(* IEC 61131-3 sources: daoli-st-library/DL_Process (part 48) *)

(* ---- FB_DL_RecipeSwitchHandover.st ---- *)
(*
  Name        : FB_DL_RecipeSwitchHandover
  Category    : DL_Process
  Version     : 1.0.0
  Purpose     : 配方切换交接编排：旧配方排空确认 → 参数装载复核（校验和整数直比）→ 新配方放行三相时序，各相独立超时故障码，中止命令相边界停下；/ Recipe switch handover orchestration: drain confirm, load recheck by integer checksum compare, release three-phase sequence with per-phase timeout fault codes and abort at phase boundary
  溯源        : 借 packml/isa88 的配方切换/批次编排组织，clean-room 实现
  Boundary    : ① 三相（排空确认/装载复核/放行）各自 TON 断输入归零 + 相超时独立锁存故障码（R40/R44）；
                ② 装载复核 = 参数集校验和整数直比，不符不放行不半装载（锁存故障至复位沿）；
                ③ 切换中收到中止命令 → 当前相边界停下（不回滚已装载段，eHold 相状态可查，信息级成因）；
                ④ 放行前复核旧配方累计量已清零反馈（幂等放行），未清零不放行（锁存故障）；
                ⑤ 命令优先级：中止 > 放行 > 装载，低优先命令直接丢弃不排队（放行仅放行相生效，装载仅空闲相受理）。
*)
TYPE E_DL_RshState :
(
    eIdle    := 0,                           (* 空闲（可受理装载命令） / Idle *)
    eDrain   := 10,                          (* 旧配方排空确认相 / Drain confirm *)
    eLoadChk := 20,                          (* 参数装载复核相 / Load recheck *)
    eRelease := 30,                          (* 新配方放行相 / Release *)
    eHold    := 40,                          (* 中止驻留相（状态可查） / Abort hold *)
    eFault   := 90                           (* 故障锁存相 / Fault latched *)
);
END_TYPE

TYPE E_DL_RshCause :
(
    eNone      := 0,                         (* 无成因 / No cause *)
    eCfgIllegal:= 1,                        (* 组态非法：相超时/周期域越界 / Illegal config *)
    eDrainTo   := 2,                        (* 排空相超时（独立码，边界①） / Drain timeout *)
    eLoadTo    := 3,                        (* 装载复核相超时（独立码） / Load recheck timeout *)
    eRelTo     := 4,                        (* 放行相超时（独立码） / Release timeout *)
    eChkMis    := 5,                        (* 校验和不符（不放行不半装载，边界②） / Checksum mismatch *)
    eAccNotClr := 6,                         (* 旧累计量未清零（不放行，边界④） / Accumulator not cleared *)
    eAbort     := 7,                        (* 中止驻留（信息级，边界③） / Abort hold, info level *)
    ePhaseBad  := 8                         (* 非法相位兜底 / Illegal phase fallback *)
);
END_TYPE

FUNCTION_BLOCK FB_DL_RecipeSwitchHandover
VAR_INPUT
    bCmdLoad : BOOL := FALSE;                (* 装载命令（仅空闲相受理，低优先丢弃）[-] / Load command *)
    bCmdRelease: BOOL := FALSE;              (* 放行命令（仅放行相复核生效）[-] / Release command *)
    bCmdAbort: BOOL := FALSE;                (* 中止命令（最高优先级，相边界停下）[-] / Abort command *)
    bDrainDone: BOOL := FALSE;               (* 排空完成反馈（属主工艺确认）[-] / Drain done feedback *)
    nChkCalc : DINT := 0;                    (* 参数集实算校验和（属主算好输入）[-] / Calculated checksum *)
    nChkExpect: DINT := 0;                   (* 期望校验和（整数直比目标）[-] / Expected checksum *)
    bAccClear: BOOL := FALSE;                (* 旧配方累计量已清零反馈 [-] / Accumulator cleared feedback *)
    tDrain   : TIME := T#30S;                (* 排空相超时，域 > T#0S [ms] / Drain phase timeout *)
    tLoadChk : TIME := T#10S;                (* 装载复核相超时 [ms] / Load phase timeout *)
    tRelease : TIME := T#5S;                 (* 放行相超时 [ms] / Release phase timeout *)
    tScan    : TIME := T#100MS;              (* 扫描周期，域 > T#0S [ms] / Scan period *)
    bEnable  : BOOL := TRUE;                 (* 使能 [-] / Enable *)
    bReset   : BOOL := FALSE;                (* 复位命令，上升沿清故障回空闲 [-] / Reset command *)
END_VAR
VAR_OUTPUT
    bReleased: BOOL;                         (* 放行完成脉冲（单拍）[-] / Released pulse *)
    bHold    : BOOL;                         (* 中止驻留指示（状态可查，边界③）[-] / Abort hold indicator *)
    nActPhase: INT;                          (* 当前生效相序号（诊断）[-] / Active phase index *)
    eState   : E_DL_RshState;                (* 状态出口 / State outlet *)
    eCause   : E_DL_RshCause;                (* 成因出口（R190 归因唯一） / Cause outlet *)
    bError   : BOOL;                         (* 故障锁存标志 [-] / Fault latch flag *)
END_VAR
VAR
    _eState : E_DL_RshState := E_DL_RshState.eIdle;  (* 内部相位（CASE 唯一写入目标） / Internal phase *)
    _eCause : E_DL_RshCause := E_DL_RshCause.eNone;  (* 成因锁存量 / Latched cause *)
    rtLoad  : R_TRIG;                        (* 装载命令沿实例，段 0 无条件调用 / Load edge instance *)
    rtReset : R_TRIG;                        (* 复位沿实例，段 0 无条件调用 / Reset edge instance *)
    tonDrain: TON;                           (* 排空相超时（IN 串相位闸，边界①） / Drain timeout *)
    tonLoadT: TON;                           (* 装载相超时（IN 串相位闸） / Load timeout *)
    tonRel  : TON;                           (* 放行相超时（IN 串相位闸） / Release timeout *)
    _bFault : BOOL;                          (* 故障锁存位 / Latched fault bit *)
    _bCfgBad: BOOL;                          (* 组态非法当拍量 / Illegal config this scan *)
    _bRelI  : BOOL;                          (* 放行脉冲内部量（统一出口映射，R187） / Release pulse internal *)
    _bChkOk : BOOL;                          (* 校验和相符当拍量（整数直比）[-] / Checksum match *)
END_VAR
VAR CONSTANT
    DL_RSH_EPS : REAL := 1.0E-6;             (* 判零容差（周期闸配套）[-] / Epsilon *)
END_VAR

(* —— 段 0：当拍判据派生 + 实例无条件刷新（R228A；TON 全段 0，边界①） —— *)
_bCfgBad := NOT (tDrain > T#0S) OR NOT (tLoadChk > T#0S) OR NOT (tRelease > T#0S) OR NOT (tScan > T#0S);   (* 相超时/周期域闸（边界①） / Timeout gates *)
rtLoad(CLK := bCmdLoad);                                 (* 装载沿每拍必调 / Load edge every scan *)
rtReset(CLK := bReset);                                  (* 复位沿每拍必调 / Reset edge every scan *)
_bChkOk := (nChkCalc = nChkExpect);                      (* 校验和整数直比（边界②） / Checksum integer compare *)
tonDrain(IN := (_eState = E_DL_RshState.eDrain), PT := tDrain);          (* 排空超时：相位闸 + 无条件调用（R40） / Drain timer *)
tonLoadT(IN := (_eState = E_DL_RshState.eLoadChk), PT := tLoadChk);      (* 装载超时：相位闸 + 无条件调用 / Load timer *)
tonRel(IN := (_eState = E_DL_RshState.eRelease), PT := tRelease);        (* 放行超时：相位闸 + 无条件调用 / Release timer *)

(* —— 段 1：单拍量预清零（R107） —— *)
_bRelI := FALSE;                                         (* 放行脉冲内部量预清 / Release preset *)
bReleased := FALSE;                                      (* 放行脉冲出口预清 / Release outlet preset *)
bHold := FALSE;                                          (* 中止指示出口预清（派生拍覆盖） / Hold preset *)
nActPhase := 0;                                          (* 相序号预清（派生拍覆盖） / Phase index preset *)

(* —— 段 2：复位沿处理（作用域：清故障 + 回空闲，R283 逐项声明） —— *)
IF rtReset.Q THEN
    _bFault := FALSE;                                    (* 清故障锁存 / Clear fault *)
    _eCause := E_DL_RshCause.eNone;                      (* 清成因 / Clear cause *)
    _eState := E_DL_RshState.eIdle;                      (* 回空闲相 / Back to idle *)
END_IF

(* —— 段 3：组态故障锁存（锁存至复位沿，R189） —— *)
IF _bCfgBad AND NOT _bFault THEN
    _bFault := TRUE;                                     (* 锁存故障位 / Latch fault *)
    _eCause := E_DL_RshCause.eCfgIllegal;                (* 成因：组态非法 / Cause illegal config *)
    _eState := E_DL_RshState.eFault;                     (* 同步迁故障相 / Migrate to fault *)
END_IF

(* —— 段 4：CASE 主状态机（ELSE 兜底迁 eFault，红线 6） —— *)
CASE _eState OF
    E_DL_RshState.eIdle:                                 (* 空闲：出口确定值，仅装载命令受理（边界⑤） / Idle *)
        IF NOT bEnable THEN
            ;                                            (* 失能保持空闲 / Disabled hold *)
        ELSIF bCmdAbort THEN
            _eCause := E_DL_RshCause.eAbort;             (* 空闲相中止：信息级记因（无相可停） / Abort in idle *)
        ELSIF rtLoad.Q AND NOT _bFault THEN              (* 装载命令沿受理（低优先级在忙相丢弃，边界⑤） / Accept load *)
            _eState := E_DL_RshState.eDrain;             (* 进入排空确认相 / Enter drain *)
        END_IF
    E_DL_RshState.eDrain:                                (* 排空确认相：反馈 or 超时 or 中止（边界①③） / Drain *)
        IF bCmdAbort THEN
            _eCause := E_DL_RshCause.eAbort;             (* 中止：信息级成因（边界③） / Abort cause *)
            _eState := E_DL_RshState.eHold;              (* 当前相边界停下（不回滚） / Hold at boundary *)
        ELSIF tonDrain.Q THEN
            _bFault := TRUE;                             (* 排空相超时独立锁存（边界①） / Drain timeout latch *)
            _eCause := E_DL_RshCause.eDrainTo;           (* 成因：排空超时 / Cause drain timeout *)
            _eState := E_DL_RshState.eFault;             (* 迁故障相 / To fault *)
        ELSIF bDrainDone THEN
            _eState := E_DL_RshState.eLoadChk;           (* 排空确认 → 装载复核相 / To load recheck *)
        END_IF
    E_DL_RshState.eLoadChk:                              (* 装载复核相：校验和直比（边界②） / Load recheck *)
        IF bCmdAbort THEN
            _eCause := E_DL_RshCause.eAbort;             (* 中止：信息级成因（边界③） / Abort cause *)
            _eState := E_DL_RshState.eHold;              (* 相边界停下 / Hold at boundary *)
        ELSIF tonLoadT.Q THEN
            _bFault := TRUE;                             (* 装载相超时独立锁存（边界①） / Load timeout latch *)
            _eCause := E_DL_RshCause.eLoadTo;            (* 成因：装载超时 / Cause load timeout *)
            _eState := E_DL_RshState.eFault;             (* 迁故障相 / To fault *)
        ELSIF NOT _bChkOk THEN
            _bFault := TRUE;                             (* 校验不符锁存：不放行不半装载（边界②） / Mismatch latch *)
            _eCause := E_DL_RshCause.eChkMis;            (* 成因：校验不符 / Cause mismatch *)
            _eState := E_DL_RshState.eFault;             (* 迁故障相（已装载段状态可查） / To fault *)
        ELSE
            _eState := E_DL_RshState.eRelease;           (* 复核通过 → 放行相 / To release *)
        END_IF
    E_DL_RshState.eRelease:                              (* 放行相：累计清零复核 + 放行命令（边界④⑤） / Release *)
        IF bCmdAbort THEN
            _eCause := E_DL_RshCause.eAbort;             (* 中止：信息级成因（边界③） / Abort cause *)
            _eState := E_DL_RshState.eHold;              (* 相边界停下 / Hold at boundary *)
        ELSIF tonRel.Q THEN
            _bFault := TRUE;                             (* 放行相超时独立锁存（边界①） / Release timeout latch *)
            _eCause := E_DL_RshCause.eRelTo;             (* 成因：放行超时 / Cause release timeout *)
            _eState := E_DL_RshState.eFault;             (* 迁故障相 / To fault *)
        ELSIF NOT bAccClear THEN
            _bFault := TRUE;                             (* 旧累计未清零不放行（幂等复核，边界④） / Acc not cleared latch *)
            _eCause := E_DL_RshCause.eAccNotClr;         (* 成因：累计未清 / Cause acc not cleared *)
            _eState := E_DL_RshState.eFault;             (* 迁故障相 / To fault *)
        ELSIF bCmdRelease THEN                           (* 放行命令在放行相生效（低优先在忙相丢弃，边界⑤） / Release command *)
            _bRelI := TRUE;                              (* 放行脉冲内部置位（R187） / Release internal *)
            _eState := E_DL_RshState.eIdle;              (* 回空闲（切换完成） / Back to idle *)
        END_IF
    E_DL_RshState.eHold:                                 (* 中止驻留相：状态可查，新装载沿重启三相（边界③） / Hold *)
        IF NOT bCmdAbort AND rtLoad.Q AND NOT _bFault THEN
            _eState := E_DL_RshState.eDrain;             (* 中止解除 + 新装载沿：从头三相（声明行为） / Restart from drain *)
        END_IF
    E_DL_RshState.eFault:                                (* 故障相：冻结保持，仅复位沿出 / Fault *)
        ;                                                (* 锁存回放（R28） / Replay from latch *)
    ELSE                                                 (* 非法相位兜底迁安全态 / Illegal phase fallback *)
        _eState := E_DL_RshState.eFault; _bFault := TRUE;    (* 迁故障相 + 同步锁存 / To fault and latch *)
        _eCause := E_DL_RshCause.ePhaseBad;              (* 成因：非法相位 / Cause illegal phase *)
END_CASE

(* —— 段 5：出口映射（内部 _b* → 输出单拍，R187；名实双出口，R191） —— *)
bReleased := _bRelI;                                     (* 放行脉冲单拍出口 / Release pulse outlet *)
bHold := (_eState = E_DL_RshState.eHold);                (* 中止驻留指示镜像 / Hold indicator mirror *)
IF _eState = E_DL_RshState.eDrain THEN
    nActPhase := 1;                                      (* 相序号：排空 / Phase drain *)
ELSIF _eState = E_DL_RshState.eLoadChk THEN
    nActPhase := 2;                                      (* 相序号：装载复核 / Phase load *)
ELSIF _eState = E_DL_RshState.eRelease THEN
    nActPhase := 3;                                      (* 相序号：放行 / Phase release *)
ELSE
    nActPhase := 0;                                      (* 空闲/驻留/故障：0（确定值） / Other phases zero *)
END_IF
bError := _bFault;                                       (* 故障标志镜像 / Fault flag mirror *)
eState := _eState;                                       (* 状态出口 / State outlet *)
eCause := _eCause;                                       (* 成因出口 / Cause outlet *)
END_FUNCTION_BLOCK

(* ---- FB_DL_ReMixerSettlerSeq.st ---- *)
(*
  Component : FB_DL_ReMixerSettlerSeq
  Category  : DL_Process
  Function  : 混合澄清槽单级串级状态机：进料→混合→澄清→（界面位越限延长分相）→排料
  Complexity: C4
  开源溯源 : DLF 内部原创（R94 族模板派生）；参考语义来源见 SOURCE_HUNTING_MATRIX.md
  规则遵从 : R1-R16
  契约     : 输入 xStart 启动（上升沿启动，下降沿兼作故障复位沿）、xStop 停止、xFeedPermit 进料许可、
             xFeedFlowOk 进料流量正常、xStageBypass 单级故障旁路、rFillPct 充液率 [%]、
             rFillTargetPct 目标充液率 [%]、rFillEmptyPct 排空判定充液率 [%]、rInterfacePct 界面位 [%]、
             rInterfHiPct 界面位上限 [%]、rInterfLoPct 界面位下限 [%]、rMixTimeS 混合时间 [s]、
             rSettleTimeS 澄清时间 [s]、rSepExtendS 分相延长时间 [s]、rFeedTmoS 进料中断超时 [s]、
             rDischTmoS 排料超时 [s]；输出五路独立命令、eState 当前相、xFault/nFaultCode 故障、
             nWarnCode 告警码、xBypassed 旁路生效、xSepExtended 处于延长分相。
  时序     : 同拍双窗配比约束 rSepExtendS ≥ rSettleTimeS（延长窗必须覆盖一个完整澄清窗，否则
             延长窗先生效、界面位尚未回稳即判超时），rFeedTmoS > 0、rDischTmoS > 0、rFillTargetPct > rFillEmptyPct。
  输出语义 : xStageBypass=TRUE 时本级输出全部撤销并停在 IDLE（不视为故障，由 xBypassed 表达）；
             xStop=TRUE 时全部命令撤销并回 IDLE（冻结保持不适用，本件为撤销型停车）。
  复位沿   : 故障码锁存至 xStart 下降沿（主路径）或 xStageBypass 上升（旁路路径），两路径均可达。
  码位     : 9810 进料许可缺失（信息级，不置 xFault）；9811 进料中断超时（故障级）；
             9812 界面位越限不可恢复（故障级）；9813 排料超时（故障级）；9814 参数或输入非法（故障级）。
*)
TYPE E_DL_ReStageState :
(
    IDLE      := 0,    // 待机，全部命令撤销 EN: idle, every command withdrawn
    FEED      := 10,   // 进料充液相 EN: feed and fill phase
    MIX       := 20,   // 混合相传质相 EN: mixing and mass transfer phase
    SETTLE    := 30,   // 澄清分相相 EN: settling and phase separation phase
    PHASE_SEP := 40,   // 界面位越限的延长分相相 EN: extended separation phase after an interface excursion
    DISCHARGE := 50,   // 排料相 EN: discharge phase
    FAULT     := 90    // 故障相，全部命令强制撤销 EN: fault phase, every command forced off
);
END_TYPE

FUNCTION_BLOCK FB_DL_ReMixerSettlerSeq
VAR_INPUT
    xStart         : BOOL;             // 启动（上升沿启动，下降沿复位故障） EN: start on the rising edge, reset the fault on the falling edge
    xStop          : BOOL;             // 停止（任意相生效，撤销全部命令） EN: stop, effective in every phase and withdrawing all commands
    xFeedPermit    : BOOL;             // 进料许可（上游供料就绪） EN: feed permit from the upstream supply
    xFeedFlowOk    : BOOL;             // 进料流量正常（流量开关） EN: the feed flow is normal, taken from the flow switch
    xStageBypass   : BOOL;             // 单级故障旁路（本级退出串级） EN: single stage fault bypass, this stage leaves the cascade
    rFillPct       : REAL;             // 槽内充液率 [%] EN: the filling level of the mixer settler
    rFillTargetPct : REAL := 85.0;     // 目标充液率（进料转混合判据） [%] EN: the target filling level that ends the feed phase
    rFillEmptyPct  : REAL := 5.0;      // 排空判定充液率 [%] EN: the filling level that ends the discharge phase
    rInterfacePct  : REAL;             // 界面位（澄清槽界面高度占比） [%] EN: the interface position as a percentage of the settler height
    rInterfHiPct   : REAL := 60.0;     // 界面位允许上限 [%] EN: the upper allowed interface position
    rInterfLoPct   : REAL := 40.0;     // 界面位允许下限 [%] EN: the lower allowed interface position
    rMixTimeS      : REAL := 300.0;    // 混合时间设定 [s] EN: the mixing time setting
    rSettleTimeS   : REAL := 600.0;    // 澄清时间设定 [s] EN: the settling time setting
    rSepExtendS    : REAL := 600.0;    // 分相延长时间设定 [s] EN: the extension time applied on an interface excursion
    rFeedTmoS      : REAL := 180.0;    // 进料中断超时设定 [s] EN: the feed interruption timeout
    rDischTmoS     : REAL := 300.0;    // 排料超时设定 [s] EN: the discharge timeout
END_VAR
VAR_OUTPUT
    xFeedValveCmd    : BOOL;               // 进料阀命令 EN: the feed valve command
    xMixerCmd        : BOOL;               // 混合搅拌命令 EN: the mixer command
    xSettlePlateCmd  : BOOL;               // 澄清挡板投入命令 EN: the settler plate command
    xDischargeCmd    : BOOL;               // 排料阀命令 EN: the discharge valve command
    eState           : E_DL_ReStageState;  // 当前相 EN: the current phase
    xFault           : BOOL;               // 故障标志（仅故障级码置位） EN: the fault flag, raised by fault class codes only
    nFaultCode       : INT;                // 故障码，锁存回放 EN: the fault code replayed from the latch
    nWarnCode        : INT;                // 告警码（9810 信息级） EN: the warning code, information class
    xBypassed        : BOOL;               // 旁路生效 EN: the bypass is active
    xSepExtended     : BOOL;               // 处于延长分相相 EN: the extended separation phase is active
    rSepElapsedS     : REAL;               // 本次分相已用时间 [s] EN: the separation time elapsed in this cycle
END_VAR
VAR
    tonFeed    : TON;                  // 进料中断超时定时器 EN: the feed interruption timeout
    tonMix     : TON;                  // 混合时间定时器 EN: the mixing timer
    tonSettle  : TON;                  // 澄清时间定时器 EN: the settling timer
    tonSep     : TON;                  // 延长分相总时间定时器 EN: the extended separation total timer
    tonDisch   : TON;                  // 排料超时定时器 EN: the discharge timeout
    fbStartRise: R_TRIG;               // xStart 上升沿（唯一启动沿） EN: the rising edge of xStart, the only start edge
    fbStartFall: F_TRIG;               // xStart 下降沿（主复位沿） EN: the falling edge of xStart, the main reset edge
    fbBypRise  : R_TRIG;               // 旁路上升沿（旁路复位路径） EN: the rising edge of the bypass, the secondary reset path
    xFinAll    : BOOL;                 // 全部浮点入参有限 EN: every floating input is finite
    xFinMix    : BOOL;                 // 混合时间有限 EN: the mixing time is finite
    xParamBad  : BOOL;                 // 参数或输入非法 EN: a parameter or an input is illegal
    xInterfOk  : BOOL;                 // 界面位在允许带内 EN: the interface position is inside the band
    xFillFull  : BOOL;                 // 充液到位 EN: the filling level reached the target
    xFillEmpty : BOOL;                 // 充液已排空 EN: the filling level dropped to the empty limit
    nMsMix     : UDINT := 300000;      // 混合毫秒数（缺省防首拍零 PT） EN: the mixing time in milliseconds, the default avoids a zero preset
    nMsSettle  : UDINT := 600000;      // 澄清毫秒数 EN: the settling time in milliseconds
    nMsSep     : UDINT := 1200000;     // 延长分相毫秒数 EN: the extended separation time in milliseconds
    nMsFeed    : UDINT := 180000;      // 进料超时毫秒数 EN: the feed timeout in milliseconds
    nMsDisch   : UDINT := 300000;      // 排料超时毫秒数 EN: the discharge timeout in milliseconds
    nCodeLatch : INT;                  // 故障码锁存副本 EN: the latched copy of the fault code
END_VAR
VAR CONSTANT
    DL_RMS_Z      : REAL := 0.0;       // 浮点零常量 EN: the floating point zero constant
    DL_RMS_K1000  : REAL := 1000.0;    // 秒转毫秒系数 EN: the second to millisecond factor
    DL_RMS_C_PERM : INT := 9810;       // 进料许可缺失（信息级） EN: the missing feed permit, information class
    DL_RMS_C_FEED : INT := 9811;       // 进料中断超时 EN: the feed interruption timeout
    DL_RMS_C_INTER: INT := 9812;       // 界面位越限不可恢复 EN: the interface excursion is not recoverable
    DL_RMS_C_DISCH: INT := 9813;       // 排料超时 EN: the discharge timeout
    DL_RMS_C_PARAM: INT := 9814;       // 参数或输入非法 EN: a parameter or an input is illegal
END_VAR

// 段1｜参数与采样门禁（先判后用：REAL→UDINT 换算在闸后执行，结果供段2 定时器 PT 使用）
xFinMix := (rMixTimeS = rMixTimeS) AND ((rMixTimeS - rMixTimeS) = DL_RMS_Z);                                     // 混合时间有限性 EN: the mixing time is finite
xFinAll := xFinMix
        AND (rFillPct = rFillPct) AND ((rFillPct - rFillPct) = DL_RMS_Z)
        AND (rFillTargetPct = rFillTargetPct) AND ((rFillTargetPct - rFillTargetPct) = DL_RMS_Z)
        AND (rFillEmptyPct = rFillEmptyPct) AND ((rFillEmptyPct - rFillEmptyPct) = DL_RMS_Z)
        AND (rInterfacePct = rInterfacePct) AND ((rInterfacePct - rInterfacePct) = DL_RMS_Z)
        AND (rInterfHiPct = rInterfHiPct) AND ((rInterfHiPct - rInterfHiPct) = DL_RMS_Z)
        AND (rInterfLoPct = rInterfLoPct) AND ((rInterfLoPct - rInterfLoPct) = DL_RMS_Z)
        AND (rSettleTimeS = rSettleTimeS) AND ((rSettleTimeS - rSettleTimeS) = DL_RMS_Z)
        AND (rSepExtendS = rSepExtendS) AND ((rSepExtendS - rSepExtendS) = DL_RMS_Z)
        AND (rFeedTmoS = rFeedTmoS) AND ((rFeedTmoS - rFeedTmoS) = DL_RMS_Z)
        AND (rDischTmoS = rDischTmoS) AND ((rDischTmoS - rDischTmoS) = DL_RMS_Z);                                 // 全部浮点入参有限性 EN: the finiteness of every floating input
xParamBad := (NOT xFinAll) OR (rMixTimeS <= DL_RMS_Z) OR (rSettleTimeS <= DL_RMS_Z) OR (rSepExtendS < DL_RMS_Z)
          OR (rFeedTmoS <= DL_RMS_Z) OR (rDischTmoS <= DL_RMS_Z)
          OR (rFillTargetPct <= rFillEmptyPct) OR (rFillEmptyPct < DL_RMS_Z)
          OR (rInterfHiPct <= rInterfLoPct);                                                                     // 域闸与配比约束 EN: the domain gate and the ratio constraints
IF NOT xParamBad THEN                                                                                            // 参数合法才做换算 EN: convert only when the parameters are legal
    nMsMix := REAL_TO_UDINT(rMixTimeS * DL_RMS_K1000);                                                           // 混合毫秒数 EN: the mixing milliseconds
    nMsSettle := REAL_TO_UDINT(rSettleTimeS * DL_RMS_K1000);                                                     // 澄清毫秒数 EN: the settling milliseconds
    nMsSep := REAL_TO_UDINT((rSettleTimeS + rSepExtendS) * DL_RMS_K1000);                                        // 延长分相毫秒数（澄清+延长） EN: the extended separation milliseconds
    nMsFeed := REAL_TO_UDINT(rFeedTmoS * DL_RMS_K1000);                                                          // 进料超时毫秒数 EN: the feed timeout milliseconds
    nMsDisch := REAL_TO_UDINT(rDischTmoS * DL_RMS_K1000);                                                        // 排料超时毫秒数 EN: the discharge timeout milliseconds
END_IF
xInterfOk := xFinAll AND (rInterfacePct <= rInterfHiPct) AND (rInterfacePct >= rInterfLoPct);                    // 界面位带内判据 EN: the interface band test
xFillFull := xFinAll AND (rFillPct >= rFillTargetPct);                                                           // 充液到位判据 EN: the fill completion test
xFillEmpty := xFinAll AND (rFillPct <= rFillEmptyPct);                                                           // 排空到位判据 EN: the empty completion test

// 段2｜五只定时器 + 三只边沿实例无条件周期刷新（R7；CASE 内不得调用实例）
tonFeed(IN := (eState = E_DL_ReStageState.FEED) AND (NOT xFeedFlowOk) AND xFeedPermit, PT := UDINT_TO_TIME(nMsFeed));  // 进料中断计时（无许可时暂停，避免关阀被误判中断） EN: time the feed interruption, paused while the permit is absent so a closed valve is not misread as an interruption
tonMix(IN := (eState = E_DL_ReStageState.MIX), PT := UDINT_TO_TIME(nMsMix));                                     // 混合计时 EN: time the mixing phase
tonSettle(IN := (eState = E_DL_ReStageState.SETTLE), PT := UDINT_TO_TIME(nMsSettle));                            // 澄清计时 EN: time the settling phase
tonSep(IN := (eState = E_DL_ReStageState.PHASE_SEP), PT := UDINT_TO_TIME(nMsSep));                               // 延长分相总计时 EN: time the extended separation phase
tonDisch(IN := (eState = E_DL_ReStageState.DISCHARGE), PT := UDINT_TO_TIME(nMsDisch));                            // 排料计时 EN: time the discharge phase
fbStartRise(CLK := xStart);                                                                                      // 启动沿 EN: the start edge
fbStartFall(CLK := xStart);                                                                                      // 复位沿 EN: the reset edge
fbBypRise(CLK := xStageBypass);                                                                                  // 旁路沿 EN: the bypass edge

// 段3｜输出预置（唯一预置点，CASE 内只置位；单拍信息位在此每拍清零）
xFeedValveCmd := FALSE;                                                                                          // 进料阀预置关 EN: preset the feed valve closed
xMixerCmd := FALSE;                                                                                              // 搅拌预置停 EN: preset the mixer off
xSettlePlateCmd := FALSE;                                                                                        // 挡板预置撤 EN: preset the settler plate withdrawn
xDischargeCmd := FALSE;                                                                                          // 排料阀预置关 EN: preset the discharge valve closed
xFault := FALSE;                                                                                                 // 故障标志预置假 EN: preset the fault flag false
nFaultCode := 0;                                                                                                 // 故障码预置零 EN: preset the fault code to zero
nWarnCode := 0;                                                                                                  // 告警码预置零 EN: preset the warning code to zero
xBypassed := xStageBypass;                                                                                       // 旁路状态直映 EN: mirror the bypass input
xSepExtended := FALSE;                                                                                           // 延长分相标志预置假 EN: preset the extension flag false
rSepElapsedS := DL_RMS_Z;                                                                                        // 分相已用时间预置零 [s] EN: preset the separation elapsed time to zero

// 段4｜全局闸：参数非法锁故障；xStop 撤销全部命令并回待机（复位沿作用域见头注释）
IF xParamBad THEN
    nCodeLatch := DL_RMS_C_PARAM;                                                                                // 参数非法锁存 EN: latch the parameter code
    xFault := TRUE;                                                                                              // 置故障标志 EN: raise the fault flag
    nFaultCode := DL_RMS_C_PARAM;                                                                                // 故障码出口 EN: publish the fault code
    eState := E_DL_ReStageState.FAULT;                                                                           // 迁故障相 EN: move to the fault phase
ELSIF xStop AND (eState <> E_DL_ReStageState.IDLE) THEN
    eState := E_DL_ReStageState.IDLE;                                                                            // 撤销型停车回待机 EN: a withdrawing stop returns to idle
END_IF

// 段5｜主状态机（ENUM + CASE，ELSE 兜底非法值）
IF eState <> E_DL_ReStageState.FAULT THEN
CASE eState OF
E_DL_ReStageState.IDLE:
    // 拍 N：待机；旁路时禁止启动（本级退出串级），启动需进料许可且无停车
    IF (NOT xStageBypass) AND fbStartRise.Q AND xFeedPermit AND (NOT xStop) AND (NOT xParamBad) THEN
        eState := E_DL_ReStageState.FEED;                                                                        // 本拍行为：进进料相 EN: enter the feed phase
    END_IF

E_DL_ReStageState.FEED:
    // 拍 N：进料充液；无许可只驻留告警（信息级），中断计时暂停，恢复许可后继续累计；有许可且中断累计超时判 9811
    // EN: feeding and filling; without the permit only an information warning is raised and the interruption timer is held, resuming when the permit returns; an interruption with the permit present raises 9811
    IF NOT xFeedPermit THEN
        nWarnCode := DL_RMS_C_PERM;                                                                              // 许可缺失告警，不置故障 EN: warn about the missing permit, no fault
    END_IF
    IF tonFeed.Q THEN
        nCodeLatch := DL_RMS_C_FEED;                                                                             // 进料中断超时 EN: the feed interruption timed out
        xFault := TRUE;                                                                                          // 置故障标志 EN: raise the fault flag
        nFaultCode := DL_RMS_C_FEED;                                                                             // 故障码出口 EN: publish the fault code
        eState := E_DL_ReStageState.FAULT;                                                                       // 迁故障相 EN: move to the fault phase
    ELSIF xFillFull THEN
        eState := E_DL_ReStageState.MIX;                                                                         // 本拍行为：进混合相 EN: enter the mixing phase
    END_IF

E_DL_ReStageState.MIX:
    // 拍 N：搅拌混合，混合时间到即转澄清
    IF tonMix.Q THEN
        eState := E_DL_ReStageState.SETTLE;                                                                      // 本拍行为：进澄清相 EN: enter the settling phase
    END_IF

E_DL_ReStageState.SETTLE:
    // 拍 N：静置澄清；界面位越限立即转延长分相，澄清时间到且界面位在带内才放行排料
    IF NOT xInterfOk THEN
        eState := E_DL_ReStageState.PHASE_SEP;                                                                   // 本拍行为：界面位越限转延长分相 EN: an interface excursion moves to the extended phase
    ELSIF tonSettle.Q AND xInterfOk THEN
        eState := E_DL_ReStageState.DISCHARGE;                                                                   // 本拍行为：澄清完成进排料相 EN: settling done, enter discharge
    END_IF

E_DL_ReStageState.PHASE_SEP:
    // 拍 N：延长分相；界面位回带内即放行，延长窗耗尽仍越限判 9812
    IF tonSep.Q AND (NOT xInterfOk) THEN
        nCodeLatch := DL_RMS_C_INTER;                                                                            // 界面位不可恢复 EN: the interface excursion is not recoverable
        xFault := TRUE;                                                                                          // 置故障标志 EN: raise the fault flag
        nFaultCode := DL_RMS_C_INTER;                                                                            // 故障码出口 EN: publish the fault code
        eState := E_DL_ReStageState.FAULT;                                                                       // 迁故障相 EN: move to the fault phase
    ELSIF xInterfOk THEN
        eState := E_DL_ReStageState.DISCHARGE;                                                                   // 本拍行为：界面位回稳进排料相 EN: the interface recovered, enter discharge
    END_IF

E_DL_ReStageState.DISCHARGE:
    // 拍 N：排料；排空回待机，排料超时判 9813（迁入本相已带参数闸复检）
    IF xParamBad THEN
        nCodeLatch := DL_RMS_C_PARAM;                                                                            // 参数退化锁存 EN: latch the parameter code
        xFault := TRUE;                                                                                          // 置故障标志 EN: raise the fault flag
        nFaultCode := DL_RMS_C_PARAM;                                                                            // 故障码出口 EN: publish the fault code
        eState := E_DL_ReStageState.FAULT;                                                                       // 迁故障相 EN: move to the fault phase
    ELSIF tonDisch.Q AND (NOT xFillEmpty) THEN
        nCodeLatch := DL_RMS_C_DISCH;                                                                            // 排料超时 EN: the discharge timed out
        xFault := TRUE;                                                                                          // 置故障标志 EN: raise the fault flag
        nFaultCode := DL_RMS_C_DISCH;                                                                            // 故障码出口 EN: publish the fault code
        eState := E_DL_ReStageState.FAULT;                                                                       // 迁故障相 EN: move to the fault phase
    ELSIF xFillEmpty THEN
        eState := E_DL_ReStageState.IDLE;                                                                        // 本拍行为：排空回待机 EN: discharged, back to idle
    END_IF

E_DL_ReStageState.FAULT:
    // 故障相（本段被外层 IF 排除，保留分支以满足枚举穷举）
    xFault := TRUE;                                                                                              // 保持故障标志 EN: keep the fault flag
    nFaultCode := nCodeLatch;                                                                                    // 锁存回放 EN: replay the latch

ELSE
    // 非法状态兜底：绝不停在未知相
    nCodeLatch := DL_RMS_C_PARAM;                                                                                // 非法状态归参数码 EN: treat an illegal state as a parameter code
    xFault := TRUE;                                                                                              // 置故障标志 EN: raise the fault flag
    nFaultCode := DL_RMS_C_PARAM;                                                                                // 故障码出口 EN: publish the fault code
    eState := E_DL_ReStageState.FAULT;                                                                           // 迁故障相 EN: move to the fault phase
END_CASE
END_IF

// 段6｜相独立使能出口（IDLE/FAULT 不置任何命令，天然强制撤销）
CASE eState OF
E_DL_ReStageState.FEED:
    xFeedValveCmd := xFeedPermit;                                                                                // 进料阀命令（无许可不投） EN: the feed valve command, gated by the permit
E_DL_ReStageState.MIX:
    xMixerCmd := TRUE;                                                                                           // 搅拌命令 EN: the mixer command
E_DL_ReStageState.SETTLE:
    xSettlePlateCmd := TRUE;                                                                                     // 澄清挡板投入 EN: the settler plate command
E_DL_ReStageState.PHASE_SEP:
    xSettlePlateCmd := TRUE;                                                                                     // 延长分相仍保持挡板 EN: the plate stays in during the extension
    xSepExtended := TRUE;                                                                                        // 延长分相标志 EN: the extension flag
    rSepElapsedS := TIME_TO_REAL(tonSep.ET) * 0.001;                                                             // 分相已用时间 [s] EN: the separation time elapsed
E_DL_ReStageState.DISCHARGE:
    xDischargeCmd := TRUE;                                                                                       // 排料阀命令 EN: the discharge valve command
ELSE
    // 其余相（含 IDLE/FAULT）：全部命令保持撤销
    xFeedValveCmd := FALSE;                                                                                      // 进料阀保持关 EN: keep the feed valve closed
    xMixerCmd := FALSE;                                                                                          // 搅拌保持停 EN: keep the mixer off
    xSettlePlateCmd := FALSE;                                                                                    // 挡板保持撤 EN: keep the plate withdrawn
    xDischargeCmd := FALSE;                                                                                      // 排料阀保持关 EN: keep the discharge valve closed
END_CASE

// 段7｜故障相锁存回放 + 两条复位路径（xStart 下降沿主路径 / 旁路上升沿旁路路径）
IF eState = E_DL_ReStageState.FAULT THEN
    xFault := TRUE;                                                                                              // 故障标志保持 EN: keep the fault flag
    nFaultCode := nCodeLatch;                                                                                    // 锁存回放，不按当下输入重推断 EN: replay the latch instead of re inferring
    nWarnCode := 0;                                                                                              // 故障相不报信息级码 EN: no information class code in the fault phase
    xFeedValveCmd := FALSE;                                                                                      // 进料阀强制关 EN: force the feed valve closed
    xMixerCmd := FALSE;                                                                                          // 搅拌强制停 EN: force the mixer off
    xSettlePlateCmd := FALSE;                                                                                    // 挡板强制撤 EN: force the plate withdrawn
    xDischargeCmd := FALSE;                                                                                      // 排料阀强制关 EN: force the discharge valve closed
    IF fbStartFall.Q OR fbBypRise.Q THEN
        nCodeLatch := 0;                                                                                         // 清除边：下降沿或旁路沿（头注释已声明） EN: clear on the falling edge or the bypass edge
        eState := E_DL_ReStageState.IDLE;                                                                        // 回待机 EN: back to idle
    END_IF
END_IF
END_FUNCTION_BLOCK

(* ---- FB_DL_RfidTrayRoute.st ---- *)
(*==============================================================================
 * 组件名称 (Component)  : FB_DL_RfidTrayRoute
 * 所属子库 (Sublibrary) : DL_Process
 * 当前版本 (Version)    : 1.0.0
 * 兼容性   (Platform)   : CODESYS 3.5+ / TwinCAT 3 / 汇川 InoProShop / 施耐德 Machine Expert
 *                         仅依赖 Standard.library（TON / R_TRIG / LEN），零厂商私有库
 * 功能描述 (Function)   : 载具 RFID 身份驱动路径路由。
 *                         读到载具身份码后在**调用者提供的路由表**中线性匹配，命中即锁定路由号并发出
 *                         段切换请求，等段间握手确认后放行；未命中则拒路由并锁存（未知载具不允许
 *                         在线上自由流动）；同一载具在防抖窗内重复读到同一码时按"重扫"忽略。
 *                         三条固化纪律：
 *                           ① **未知载具拒路由**：匹配失败即锁存 bUnknownTray 并进故障相，
 *                              绝不给"默认路由"兜底（默认路由会把未知载具送进错误工位）；
 *                           ② **重复读码防抖**：路由成功后置防抖窗（tDupWin），窗内读到**同一码**
 *                              只置 bDupRead（信息级），不改路由、不重发段请求；读到**不同码**
 *                              视为换载具，立即重匹配；
 *                           ③ **段间握手**：请求脉冲单拍、等确认超时锁存，超时与不一致分码归因。
 *                         验收向量：
 *                           ① 路由表 3 条 {TRAY-A, TRAY-B, TRAY-C}，读 TRAY-B → iRouteNo = 2
 *                           ② 读 TRAY-Z → 拒路由 + bUnknownTray 锁存（等复位）
 *                           ③ 读 TRAY-B 后 tDupWin 内再读 TRAY-B → bDupRead 单拍，iRouteNo 不变
 *                           ④ 段请求发出后超时无 bSegAck → bUnknownTray 不动，锁存 eSegTimeout
 * 接口     (Interface)  : 入 bReadDone 读码完成沿、sTrayId 载具身份码、bStartSeg 段切换启动沿、
 *                         bSegAck 段间确认、nRouteCnt 路由表有效条数、tDupWin 防抖窗、
 *                         tSegAckTo 段握手超时、bReset 复位沿；
 *                         路由表 IN_OUT asRouteTable（1..16，调用者持有）；
 *                         出 iRouteNo 路由号（0 = 无）、bRouteValid 路由就绪、bSegReq 段请求脉冲（单拍）、
 *                         bSegBusy 等确认中、bUnknownTray 未知载具锁存、bDupRead 重扫忽略脉冲（单拍）、
 *                         eState 相、eCause 成因、bError 故障标志。
 * 边界     (Boundary)   : ① **属主边界（写死）：本件只做"身份 → 路由号 → 段放行"，
 *                         不驱动读码头、不驱动输送段电机、不写 MES 履历**；
 *                         ② **路由表边界**：表上界以字面量 16 声明（R104），有效条数 nRouteCnt 作
 *                         运行时二次闸（钳 0..16）；匹配循环带 _uGuard 计数，必然收敛；
 *                         ③ **空码闸**：LEN(sTrayId) = 0 → 视为无码，拒路由 + eNoCode（信息级，不锁存）；
 *                         ④ **超时 TON 冻结**：tonSeg / tonDup 的 IN 均串 (NOT _bFault)，
 *                         故障期不累计，复位同拍不会立即重锁（R252）；
 *                         ⑤ **锁存解除式**：bUnknownTray 与 eFault 仅由 bReset 上升沿解除
 *                         （R228B 唯一迁出）；bReset 为外部引脚，恒可达；
 *                         ⑥ 零全局耦合、零物理地址。
 * 分工声明 (Scope)      : 本件只管"载具身份路由编排"。不接管：读码头驱动与标签数据块解析
 *                         （属 FB_DL_RfidTagHandler 族）、FOUP 配方放行校验（属 FB_DL_FoupRfidCheck）、
 *                         输送段方向控制（属输送件）。
 * 来源标签 (Source Tag) : ROADMAP 空勾真缺口 P1（RFID 载具路由，自研 clean-room）
 * 码表     (Codes)      : 本件不占用任何全局数字码位（零码位范式 R297）；诊断由 BOOL + ENUM 出口承担。
 * 红线自检 (Redline)    : R1 ✓ 零 GVL/VAR_EXTERNAL ｜ R2 ✓ 零 %I/%Q/%M ｜ R3 ✓ 纯 IEC 61131-3
 *                         R4 ✓ 表界闸 + 循环计数器 + 空码闸 + 双超时 ｜ R5 ✓ 声明逐行同行双语注释
 *                         R6 ✓ ENUM+CASE 含 ELSE 兜底 ｜ R7 ✓ 双 TON/三 R_TRIG 段 0 无条件刷新
 * 修订历史 (Revision)   : 2026-11-19  v1.0.0  R47 首版（批次 3 · 序号 11）
 *==============================================================================*)

TYPE E_DL_RtrState :
(
    eIdle   := 0,    // 待机相（等读码） / Idle, awaiting a tag read
    eSegWait:= 10,   // 等段确认相（握手窗口内） / Waiting for the segment acknowledgement
    eFault  := 90    // 故障相（等复位） / Fault, awaiting reset
);
END_TYPE

TYPE E_DL_RtrCause :
(
    eNone      := 0,   // 无异常 / No anomaly
    eUnknownTray:= 1,  // 未知载具（拒路由，锁存） / Unknown tray, routing refused, latched
    eNoCode    := 2,   // 空码（信息级，不锁存） / Empty code, info level
    eDupRead   := 3,   // 防抖窗内重扫（信息级，不锁存） / Duplicate read inside the debounce window
    eSegTimeout:= 4,   // 段握手超时（锁存） / Segment handshake timeout, latched
    eCfgIllegal:= 5,   // 组态非法（路由表条数/时间越域） / Illegal configuration
    ePhaseBad  := 6    // 非法相位兜底 / Illegal phase fallback
);
END_TYPE

FUNCTION_BLOCK FB_DL_RfidTrayRoute
VAR_IN_OUT
    asRouteTable : ARRAY[1..16] OF STRING[15];   // 路由表（1..16，条内容由调用者维护） [-] / Route table owned by the caller
END_VAR
VAR_INPUT
    bReadDone  : BOOL := FALSE;      // 读码完成沿 [-] / Tag-read edge
    sTrayId    : STRING[15] := '';   // 载具身份码（≤15 字符） [-] / Tray identity code
    bStartSeg  : BOOL := FALSE;      // 段切换启动沿 [-] / Segment-start edge
    bSegAck    : BOOL := FALSE;      // 段间确认（当拍电平） [-] / Segment acknowledgement, level
    nRouteCnt  : INT := 0;           // 路由表有效条数，域 0..16 [条] / Valid route count, 0..16
    tDupWin    : TIME := T#5S;       // 重复读码防抖窗，域 > T#0S [ms] / Duplicate-read debounce window
    tSegAckTo  : TIME := T#10S;      // 段握手超时，域 > T#0S [ms] / Segment handshake timeout
    bReset     : BOOL := FALSE;      // 故障复位沿 [-] / Fault reset edge
END_VAR
VAR_OUTPUT
    iRouteNo    : INT := 0;                              // 路由号（1..16；0 = 无） [-] / Route number, 0 = none
    bRouteValid : BOOL := FALSE;                         // 路由就绪（等段启动） [-] / Route ready
    bSegReq     : BOOL := FALSE;                         // 段请求脉冲（单拍） [-] / Segment request, single scan
    bSegBusy    : BOOL := FALSE;                         // 等段确认中 [-] / Waiting for the acknowledgement
    bUnknownTray: BOOL := FALSE;                         // 未知载具锁存（等复位） [-] / Unknown tray, latched
    bDupRead    : BOOL := FALSE;                         // 重扫忽略脉冲（单拍） [-] / Duplicate-read pulse
    eState      : E_DL_RtrState := E_DL_RtrState.eIdle;  // 相出口 [-] / Phase outlet
    eCause      : E_DL_RtrCause := E_DL_RtrCause.eNone;  // 成因出口（R190 归因唯一） [-] / Cause outlet
    bError      : BOOL := FALSE;                         // 故障标志（仅故障级成因） [-] / Error flag, fault level only
END_VAR
VAR
    _eState   : E_DL_RtrState := E_DL_RtrState.eIdle;    // 内部相（CASE 唯一写入目标） / Internal phase
    _eCause   : E_DL_RtrCause := E_DL_RtrCause.eNone;    // 成因锁存量 / Latched cause
    _bFault   : BOOL := FALSE;                           // 故障锁存位 / Latched fault bit
    _bUnknown : BOOL := FALSE;                           // 未知载具锁存位 / Latched unknown-tray bit
    _iRoute   : INT := 0;                                // 内部路由号 / Internal route number
    _iCnt     : INT := 0;                                // 归一后的有效条数 / Normalised valid count
    _iIdx     : INT := 0;                                // 匹配下标（1..16） / Match index
    _iHitIdx  : INT := 0;                                // 首个命中号（0 = 未命中） / First hit index, 0 = no hit
    _uGuard   : UINT := 0;                               // 匹配循环计数器（防死循环） / Match-loop guard
    _bHit     : BOOL := FALSE;                           // 匹配命中标志 / Match-found flag
    _bSegReq  : BOOL := FALSE;                           // 段请求脉冲内部位（单拍） / Internal segment request
    _bDupRead : BOOL := FALSE;                           // 重扫脉冲内部位（单拍） / Internal duplicate pulse
    _bDupBlk  : BOOL := FALSE;                           // 防抖窗封锁位（持窗量） / Debounce window blocking bit
    _sLastId  : STRING[15] := '';                        // 上次成功路由的身份码 / Last successfully routed identity
    _bCfgBad  : BOOL := FALSE;                           // 组态非法当拍量 / Illegal configuration this scan
    tonSeg    : TON;                                     // 段握手超时实例，段 0 无条件调用 / Segment timeout instance
    tonDup    : TON;                                     // 防抖窗实例，段 0 无条件调用 / Debounce window instance
    rtRead    : R_TRIG;                                  // 读码沿实例，段 0 无条件调用 / Tag-read edge instance
    rtStartSeg: R_TRIG;                                  // 段启动沿实例，段 0 无条件调用 / Segment-start edge instance
    rtReset   : R_TRIG;                                  // 复位沿实例，段 0 无条件调用 / Reset edge instance
END_VAR
VAR CONSTANT
    DL_RTR_MAX   : INT := 16;            // 路由表深度（与数组字面量上界同源） [条] / Route table depth
    DL_RTR_GUARD : UINT := 18;           // 匹配循环守护上限（深度 + 2） [次] / Match-loop guard limit
END_VAR

(* —— 段 0：组态闸 + 双 TON 与三沿无条件周期刷新（R228A；IN 串故障否决，R252） —— *)
_bCfgBad := (nRouteCnt < 0) OR (nRouteCnt > DL_RTR_MAX)              // 条数须在 0..16 / Count within 0..16
         OR (tDupWin <= T#0S) OR (tSegAckTo <= T#0S);                // 两时间须为正 / Both times positive
rtRead(CLK := bReadDone);                                            // 读码沿 / Tag-read edge
rtStartSeg(CLK := bStartSeg);                                        // 段启动沿 / Segment-start edge
rtReset(CLK := bReset);                                              // 复位沿 / Reset edge
tonDup(IN := _bDupBlk AND (NOT tonDup.Q), PT := tDupWin);             // 防抖窗（自复位振荡，R188） / Debounce window, self-resetting
tonSeg(IN := (_eState = E_DL_RtrState.eSegWait) AND (NOT _bFault), PT := tSegAckTo);   // 段握手超时 / Segment handshake timeout

(* —— 段 1：单拍量预清零（锁存量 _eCause/_bFault/_bUnknown/_iRoute/_bDupBlk 不入清单，R107） —— *)
bRouteValid := FALSE;                                                // 路由就绪预清 / Route-ready preset
bSegReq     := FALSE;                                                // 段请求预清（出口侧，段 6 由内部位覆写） / Segment request preset
_bSegReq    := FALSE;                                                // 段请求内部位预清 / Internal segment request preset
_bDupRead   := FALSE;                                                // 重扫脉冲内部位预清 / Internal duplicate pulse preset
bError      := FALSE;                                                // 故障标志预清（R45 配对） / Error preset

(* —— 段 2：组态闸（非法即锁存故障级） —— *)
IF _bCfgBad THEN
    _eCause := E_DL_RtrCause.eCfgIllegal;                            // 归因：组态非法 / Cause: illegal configuration
    _bFault := TRUE;                                                 // 锁存 / Latch
    _eState := E_DL_RtrState.eFault;                                 // 入故障相 / Enter fault phase
END_IF

(* —— 段 3：迁出链（bReset 上升沿：清双锁存与路由号，R228B） —— *)
IF rtReset.Q THEN
    _bFault   := FALSE;                                              // 清故障锁存 / Clear fault latch
    _bUnknown := FALSE;                                              // 清未知载具锁存 / Clear the unknown-tray latch
    _eCause   := E_DL_RtrCause.eNone;                                // 清成因 / Clear cause
    _iRoute   := 0;                                                  // 路由号清零 / Route number cleared
    _bDupBlk  := FALSE;                                              // 解除防抖封锁 / Release the debounce block
    _sLastId  := '';                                                 // 清上次身份码 / Clear the last identity
    _eState   := E_DL_RtrState.eIdle;                                // 回待机相 / Back to idle
END_IF

(* —— 段 4：防抖窗到时自动解除封锁（持窗量，非每拍预清零量） —— *)
IF tonDup.Q THEN
    _bDupBlk := FALSE;                                               // 窗到：解除封锁 / Window elapsed, release
END_IF

(* —— 段 5：读码与匹配（未知载具拒路由；同一码防抖忽略） —— *)
_iCnt := nRouteCnt;                                                  // 归一有效条数 / Normalise the valid count
IF _iCnt > DL_RTR_MAX THEN
    _iCnt := DL_RTR_MAX;                                             // 二次上界钳 / Second upper clamp
END_IF

IF (rtRead.Q) AND (NOT _bFault) AND (NOT _bCfgBad) THEN
    IF LEN(sTrayId) = 0 THEN
        _eCause := E_DL_RtrCause.eNoCode;                            // 归因：空码（信息级） / Cause: empty code, info level
    ELSIF _bDupBlk AND (sTrayId = _sLastId) THEN
        _bDupRead := TRUE;                                           // 防抖窗内同一码：重扫忽略 / Same code inside the window: ignored
        _eCause := E_DL_RtrCause.eDupRead;                           // 归因：重扫（信息级） / Cause: duplicate read, info level
    ELSE
        (* 线性匹配（带守护计数；仅记录首个命中号，未命中即非法载具） *)
        _bHit    := FALSE;                                           // 命中标志预置 / Hit preset
        _uGuard  := 0;                                               // 守护计数归零 / Guard reset
        _iIdx    := 1;                                               // 从表首匹配 / Start at the table head
        _iHitIdx := 0;                                               // 命中号预置 / Hit index preset
        WHILE (_uGuard < DL_RTR_GUARD) AND (_iIdx <= _iCnt) DO
            IF (NOT _bHit) AND (asRouteTable[_iIdx] = sTrayId) THEN
                _bHit    := TRUE;                                    // 首个命中即锁定 / Lock on the first hit
                _iHitIdx := _iIdx;                                   // 记录命中号 / Record the hit index
            END_IF
            _uGuard := _uGuard + 1;                                  // 计数器推进 / Guard advance
            _iIdx   := _iIdx + 1;                                    // 下标推进 / Index advance
        END_WHILE

        IF _bHit THEN
            _iRoute  := _iHitIdx;                                    // 锁定路由号 / Lock the route number
            _sLastId := sTrayId;                                     // 记录身份码 / Remember the identity
            _bDupBlk := TRUE;                                        // 开防抖窗 / Open the debounce window
            bRouteValid := TRUE;                                     // 路由就绪 / Route ready
        ELSE
            _bUnknown := TRUE;                                       // 未知载具：锁存 / Unknown tray: latch
            _bFault   := TRUE;                                       // 故障锁存 / Latch the fault
            _eCause   := E_DL_RtrCause.eUnknownTray;                 // 归因：未知载具 / Cause: unknown tray
            _eState   := E_DL_RtrState.eFault;                       // 入故障相 / Enter fault phase
            _iRoute   := 0;                                          // 路由号清零（拒路由） / Route number cleared
        END_IF
    END_IF
END_IF

(* —— 段 6：相迁移（段握手闭环） —— *)
IF (NOT _bFault) AND (NOT _bCfgBad) THEN
    CASE _eState OF

    E_DL_RtrState.eIdle:
        IF rtStartSeg.Q AND (_iRoute > 0) THEN
            _bSegReq := TRUE;                                        // 段请求脉冲（内部位） / Internal segment request
            _eState  := E_DL_RtrState.eSegWait;                      // 进等确认相 / Enter the wait-ack phase
        END_IF

    E_DL_RtrState.eSegWait:
        IF bSegAck THEN
            _iRoute := 0;                                            // 确认到达：路由消费完毕 / Acknowledged, the route is consumed
            _eState := E_DL_RtrState.eIdle;                          // 回待机相 / Back to idle
        ELSIF tonSeg.Q THEN
            _bFault := TRUE;                                         // 握手超时：锁存 / Timeout: latch
            _eCause := E_DL_RtrCause.eSegTimeout;                    // 归因：段握手超时 / Cause: segment timeout
            _eState := E_DL_RtrState.eFault;                         // 入故障相 / Enter fault phase
        END_IF

    E_DL_RtrState.eFault:
        ;                                                            // 故障相：仅等复位沿 / Wait for the reset edge only

    ELSE
        _eCause := E_DL_RtrCause.ePhaseBad;                          // 归因：非法相位 / Cause: illegal phase
        _bFault := TRUE;                                             // 锁存 / Latch
        _eState := E_DL_RtrState.eFault;                             // 强拉故障相 / Force fault phase

    END_CASE
END_IF

(* —— 段 7：出口单点映射（名实双出口，R191） —— *)
bSegReq     := _bSegReq;                                             // 段请求脉冲出口 / Segment request outlet
bDupRead    := _bDupRead;                                            // 重扫脉冲出口 / Duplicate-read outlet
iRouteNo    := _iRoute;                                              // 路由号出口 / Route number outlet
bSegBusy    := (_eState = E_DL_RtrState.eSegWait);                   // 等确认中出口 / Busy outlet
bUnknownTray:= _bUnknown;                                            // 未知载具出口 / Unknown-tray outlet
eState      := _eState;                                              // 相出口 / Phase outlet
eCause      := _eCause;                                              // 成因出口 / Cause outlet
bError      := _bFault;                                              // 故障标志 / Error flag

END_FUNCTION_BLOCK

(* ---- FB_DL_RfReflectedMonitor.st ---- *)
(*
  FB_DL_RfReflectedMonitor  —  射频正反功率比监视与匹配器联动告警 / RF forward-reflected power ratio monitor
  分类 Category : DL_Process
  码位 Code     : 16#06_0_B3
  版本 Version  : 1.0.0
  来源 Source   : t2-1-lgf-measurement — IEC 61131-3 标准语义的道莅防御性实现
  溯源 Origin   : clean-room 实现，射频反射比监视公开语义借鉴，未复制任何源码行（RESUME 承接 R36 §4 #18 规格）
                  （仅监视件：本件只做比值判级与请求置位，不闭环调谐——闭环调谐由匹配器本体承载，此语义为规格强制）
  功能 Function : 1) 反射比 = 反射/正向 × 100，两级阈值（Warn/Fault）带迟滞与去抖；
                  2) bMatcherRequest 在越 Warn 阈时置位并持续 tMatcherReqHold（仅请求，不闭环）；
                  3) 比值 > 100%（反射 > 正向）属异常物理值，钳到 100 并置码。
  边界 Boundary : ① fPowerFwdW <= 0 时比值不计算（防除零），输出 0 并置「无正向功率」信息码；
                  ② 组态非法（Warn >= Fault / 阈值 <= 0 / 去抖 <= 0）判组态错；
                  ③ 信号非有限（NaN 用 x<>x 自反）判无效置码，判级维持安全缺省；
                  ④ bReflFault 解除式自证：比值回落到 Warn 阈以下 AND bReset（两引脚可满足）；
                  ⑤ 本件无状态机 ENUM/CASE（监视件），判级为去抖+锁存量承载，每拍出口单点映射。
  依赖 Depends  : 仅 Standard.library（TON/TOF/ABS）；语义对齐 FB_DL_SignalStatistics / FB_DL_ToleranceWindow（已注册，不实例化）
  码表 Error codes（本件格 06_0_B3，子码步进 +0x100）:
    16#0006_01B3 信息级：无正向功率，比值不计算
    16#0006_02B3 故障级：组态非法（阈值域倒置 / 去抖 <= 0），每拍重申
    16#0006_03B3 信息级：反射功率超正向（物理异常），比值钳 100
    16#0006_04B3 信息级：匹配器请求挂起（仅请求不闭环）
    16#0006_05B3 故障级：反射比越故障阈（去抖确认，锁存至复位 + 回落）

  修订历史 Revision :
    2026-11-18  v1.0.0  R38 首版
*)

FUNCTION_BLOCK FB_DL_RfReflectedMonitor
VAR_INPUT
    fPowerFwdW       : REAL := 100.0;   // 正向功率 [W] / Forward power
    fPowerReflW      : REAL := 0.0;     // 反射功率 [W] / Reflected power
    fReflRatioWarnPct: REAL := 10.0;    // 反射比预警阈 [%] / Reflected ratio warn threshold
    fReflRatioFaultPct: REAL := 20.0;   // 反射比故障阈 [%] / Reflected ratio fault threshold
    tRatioDebounce   : TIME := T#1S;    // 判级去抖 [ms]，域 > 0 / Ratio debounce
    tMatcherReqHold  : TIME := T#30S;   // 匹配器请求保持 [ms] / Matcher request hold
    bReset           : BOOL := FALSE;   // 复位（故障锁存解除路径之一）/ Reset
END_VAR
VAR_OUTPUT
    fReflRatioPct    : REAL;            // 反射比 [%] / Reflected ratio
    bReflWarn        : BOOL;            // 预警级判级 / Warn verdict
    bReflFault       : BOOL;            // 故障级判级锁存 / Fault verdict latch
    bMatcherRequest  : BOOL;            // 匹配器请求（仅请求不闭环）/ Matcher request, monitor-only
    nErrId           : UDINT;           // 事件码，0 = 无事件 / Event code
END_VAR
VAR
    tonWarnDly  : TON;                   // 预警级去抖计时，段 0 无条件刷新 / Warn debounce timer
    tonFaultDly : TON;                   // 故障级去抖计时，段 0 无条件刷新 / Fault debounce timer
    tofReqHold  : TOF;                   // 匹配器请求保持（TOF 断输入延时），段 0 无条件刷新 / Request hold, falling-delay
    tonFaultWch : TON;                   // 故障观察窗，自复位 / Fault watch window, self-resetting
    rtReset     : R_TRIG;                // 复位上升沿 / Reset rising edge
    _rRatio     : REAL;                  // 比值暂存 [%] / Ratio scratch
    _bFwdOk     : BOOL;                  // 正向功率有效标志 / Forward power validity flag
    _bFin       : BOOL;                  // 非有限筛查标志 / Non-finite screening flag
    _bFaultL    : BOOL;                  // 故障级锁存保持量 / Fault verdict latch
    _bCfgBad    : BOOL;                  // 组态非法聚合 / Configuration invalid aggregate
    _uInfo      : UDINT;                 // 信息码，每拍重算 / Info code
END_VAR
VAR CONSTANT
    DL_WATCH_PT : TIME := T#2S;   // 故障观察窗 [ms]，自复位 / Fault watch window
END_VAR

(* —— 段 0：定时器与边沿无条件周期刷新（R182：调用语句不得置于 IF/CASE 内） —— *)
rtReset(CLK := bReset);                                          // 复位上升沿，每拍必调
tonFaultWch(IN := (NOT tonFaultWch.Q), PT := DL_WATCH_PT);       // 观察窗自复位（表达式入参）
tonWarnDly(IN := (_rRatio > fReflRatioWarnPct) AND (NOT _bCfgBad), PT := tRatioDebounce);   // 预警去抖（表达式入参）
tonFaultDly(IN := (_rRatio > fReflRatioFaultPct) AND (NOT _bCfgBad), PT := tRatioDebounce); // 故障去抖（表达式入参）
tofReqHold(IN := (_rRatio > fReflRatioWarnPct) AND (NOT _bCfgBad) AND (NOT _bFaultL),
           PT := tMatcherReqHold);                               // 请求保持（TOF，表达式入参）

(* —— 段 1：单拍量预清零（锁存量 _bFaultL 不入清单，R187①） —— *)
_uInfo := 16#0000_0000;              // 信息码每拍重算
bReflWarn := FALSE;                  // 预警出口缺省 FALSE（段 6 单点置位）
_bCfgBad := FALSE;                   // 组态非法预清零
nErrId := 16#0000_0000;              // 事件码缺省无事件

(* —— 段 2：组态域闸（覆盖全部参与判据换算的引脚，R151） —— *)
IF (fReflRatioWarnPct <= 0.0) OR (fReflRatioFaultPct <= fReflRatioWarnPct)
   OR (TIME_TO_DINT(tRatioDebounce) <= 0) THEN
    _bCfgBad := TRUE;                // 阈值域倒置或去抖非法
    nErrId := 16#0006_02B3;          // 故障级：组态非法（每拍重申）
END_IF

(* —— 段 3：信号有效性与比值计算（防除零 + 非有限筛查） —— *)
_bFin := (fPowerFwdW = fPowerFwdW) AND (fPowerReflW = fPowerReflW)
         AND (ABS(fPowerFwdW) < 1.0E15) AND (ABS(fPowerReflW) < 1.0E15);   // NaN 用 x<>x 自反
IF (NOT _bFin) OR (fPowerFwdW <= 0.0) THEN
    _bFwdOk := FALSE;                // 正向功率无效：比值不计算（防除零，规格强制）
    _rRatio := 0.0;                  // 输出 0
    IF fPowerFwdW <= 0.0 THEN
        _uInfo := 16#0006_01B3;      // 信息级：无正向功率
    END_IF
ELSE
    _bFwdOk := TRUE;                 // 分母有效
    IF fPowerReflW > fPowerFwdW THEN
        _rRatio := 100.0;            // 反射 > 正向：异常物理值钳 100（规格强制）
        _uInfo := 16#0006_03B3;      // 信息级：物理异常已钳制
    ELSE
        _rRatio := fPowerReflW * 100.0 / fPowerFwdW;   // 反射比 [%]（分母已闸 > 0）
    END_IF
END_IF
fReflRatioPct := _rRatio;            // 比值出口

(* —— 段 4：判级与锁存（故障级锁存至复位 + 回落，解除式自证） —— *)
IF _bFwdOk AND (NOT _bCfgBad) THEN
    IF tonFaultDly.Q THEN
        _bFaultL := TRUE;            // 故障级锁存（去抖确认）
    END_IF
    IF _bFaultL THEN
        IF (_rRatio <= fReflRatioWarnPct) AND rtReset.Q THEN
            _bFaultL := FALSE;       // 解除式自证：比值回落至 Warn 阈以下 AND bReset
        END_IF
    END_IF
END_IF

(* —— 段 5：出口单点映射（名实同源；锁存码回放，禁同拍抹除） —— *)
bReflFault := _bFaultL;              // 故障级出口 = 锁存量（置位同拍不被抹）
bReflWarn := tonWarnDly.Q AND (NOT _bFaultL);   // 预警出口（去抖确认，故障级优先）
bMatcherRequest := tofReqHold.Q AND (NOT _bCfgBad);   // 匹配器请求（仅请求不闭环，TOF 保持）
IF bMatcherRequest THEN
    _uInfo := 16#0006_04B3;          // 信息级：请求挂起
END_IF
IF _bCfgBad THEN
    bReflWarn := FALSE;              // 组态错判级出口撤销（安全侧）
    bMatcherRequest := FALSE;
    bReflFault := FALSE;
END_IF
IF (NOT _bCfgBad) THEN
    IF bReflFault THEN
        nErrId := 16#0006_05B3;      // 故障级码回放（锁存）
    ELSIF _uInfo <> 16#0000_0000 THEN
        nErrId := _uInfo;            // 信息码
    END_IF
END_IF

END_FUNCTION_BLOCK

(* ---- FB_DL_RollChangeoverSeq.st ---- *)
(*
  Component : FB_DL_RollChangeoverSeq
  Category  : DL_Process
  Type      : FB
  Version   : 1.0.1
  CodeSeg   : 16#06_0_3F
  Summary   : 换卷换规格一键切换顺控：参数配方合法性校验（首失败项索引）+ 张力回零超时守护 + 步进状态机。
              Roll changeover sequence: recipe validation with first-fail index plus tension zeroing timeout and step machine.
  溯源声明  : 仅借 t2-isa88 换卷流程分类与步序域，代码 clean-room（T2 借鉴件）
  边界安全  : 配方参数域闸逐项校验并输出首失败项索引（拒绝启动，按派单要点）；
              张力回零判据带超时（tZeroMs 输入引脚），不得无限等待；步进 CASE 必带 ELSE 安全步；
              张力零位判据带容差（禁等值直比）；故障码锁存有复位沿可达解除路径；TON 每拍无条件刷新。
  复用      : 复用 FB_DL_StepSequencer + FB_DL_InterlockMatrix 语义（clean-room 自含实现，无实例依赖）
*)

FUNCTION_BLOCK FB_DL_RollChangeoverSeq
VAR_INPUT
    bRun        : BOOL;                 (* 顺控使能 · Enable *)
    bStartCmd   : BOOL;                 (* 一键切换指令 [事件]，沿触发 · One-key start command *)
    fTenNowN    : LREAL;                (* 当前张力反馈 [N] · Current tension feedback *)
    fTensionSetN: LREAL := 50.0;        (* 配方：新卷张力给定 [N] · Recipe tension setpoint *)
    fSpdMpm     : LREAL := 120.0;       (* 配方：新规格线速 [m/min] · Recipe line speed *)
    fSpdMaxMpm  : LREAL := 300.0;       (* 线速上限 [m/min] · Speed upper bound *)
    fTenMaxN    : LREAL := 120.0;       (* 张力上限 [N] · Tension upper bound *)
    fZeroEpsN   : LREAL := 1.0;         (* 张力零位判据容差 [N] · Tension zero tolerance *)
    tZeroMs     : TIME  := T#8000MS;    (* 张力回零超时 [ms] · Tension zeroing timeout *)
    bReset      : BOOL;                 (* 故障复位 [事件]，沿触发 · Fault reset, edge *)
    fEps        : LREAL := 1.0E-6;      (* 浮点判零容差 [实数域] · Floating zero tolerance *)
END_VAR
VAR_OUTPUT
    eStep    : (eStpIdle := 0, eStpValidate := 1, eStpTenZero := 2, eStpSwitch := 3);   (* 步枚举输出 / Step output enum *)
    nFailIdx : INT;                     (* 配方首失败项索引 [索引]，0 为全过 · First failed recipe index *)
    bRejected: BOOL;                    (* 配方拒绝启动标志 · Recipe rejected flag *)
    bSeqDone : BOOL;                    (* 切换完成脉冲 [脉冲] · Changeover done pulse *)
    bError   : BOOL;                    (* 故障标志，与故障码配对 · Fault flag paired with codes *)
    uErrorId : UDINT;                   (* 事件码 16#0000_003F，0 无事件 · Event code *)
END_VAR
VAR
    _bDone   : BOOL;                   (* 完成脉冲内部标志 [开关] · Internal done flag *)
    _eState  : (eStIdle := 0, eStValidate := 1, eStTenZero := 2, eStSwitch := 3);   (* 内部步进状态 / Internal step state *)
    uCode    : WORD;    (* 码位暂存（锁存），复位沿清 [码] · Latched code staging *)
    tonZero  : TON;     (* 张力回零超时计时 [ms]，每拍无条件刷新 · Zeroing timeout timer *)
    rTrigStrt: R_TRIG;  (* 起动沿检测 · Start edge *)
    rTrigRst : R_TRIG;  (* 复位沿检测 · Reset edge *)
    bSigOk   : BOOL;    (* 输入有效标志 · Input validity flag *)
    nCycles  : UDINT;   (* 完成切换计数 [次]，防回卷 · Changeover count *)
END_VAR
VAR CONSTANT
    DL_RCS_WRAP : UDINT := 4294967290;  (* 计数防回卷余量 [次] · Counter wrap guard *)
END_VAR

(* === 段 0 · 实例刷新（每拍无条件，红线 7）=== *)
tonZero(IN := (_eState = eStTenZero), PT := tZeroMs);   (* 回零超时计时 / Zeroing timeout *)
rTrigStrt(CLK := bStartCmd);                            (* 起动沿检测 / Start edge *)
rTrigRst(CLK := bReset);                                (* 复位沿检测 / Reset edge *)

(* === 段 1 · 输入校验与量程闸 === *)
bSigOk := (fTenNowN = fTenNowN) AND (ABS(fTenNowN) < 1.0E308)       // 非有限拦截 / Non-finite guard
          AND (tZeroMs > T#0MS) AND (fZeroEpsN > fEps)               // 超时/容差正域闸 / Timeout and tolerance gates
          AND (fSpdMaxMpm > fEps) AND (fTenMaxN > fEps);             // 上限正域闸 / Upper bound gates
IF rTrigRst.Q THEN
    uCode := 16#0000;                   (* 复位沿清锁存（可达解除路径）/ Reset edge clears the latch *)
END_IF

(* === 段 2 · 主逻辑：配方校验与步进状态机 === *)
CASE _eState OF
    eStIdle:                            (* 空闲步：待令 / Idle *)
        IF bRun AND bSigOk AND rTrigStrt.Q THEN
            nFailIdx := 0;              (* 启动沿才清失败项，拒绝结果保留到下次启动 / Clear only on start edge *)
            bRejected := FALSE;         (* 启动沿清拒绝标志 / Clear reject on start edge *)
            uCode := 16#0000;           (* 启动沿清历史锁存码（可达解除路径 2）/ Clear latched codes on start *)
    _eState := eStValidate;     (* 拍 N 起动沿进入，拍 N+1 校验步 / To validate *)
        END_IF
    eStValidate:                        (* 校验步：逐项域闸，记首失败项 / Validate recipe, record first fail *)
        nFailIdx := 0;                  (* 默认全过 / Default all pass *)
        IF (fTensionSetN <= fEps) OR (fTensionSetN > fTenMaxN) THEN
            nFailIdx := 1;              (* 首失败项 1：张力给定域外 / Fail index 1: tension *)
        ELSIF (fSpdMpm <= fEps) OR (fSpdMpm > fSpdMaxMpm) THEN
            nFailIdx := 2;              (* 首失败项 2：线速域外 / Fail index 2: speed *)
        END_IF
        IF nFailIdx > 0 THEN
            bRejected := TRUE;          (* 拒绝启动并上报首失败项 / Reject with the first fail index *)
            uCode := 16#003F;           (* 故障级：配方域外 / Fault: recipe out of domain *)
            _eState := eStIdle;         (* 回空闲安全步 / Back to idle *)
        ELSE
            _eState := eStTenZero;      (* 校验通过转张力回零步 / To tension zeroing *)
        END_IF
    eStTenZero:                         (* 回零步：张力进入零位容差带 / Zeroing with tolerance band *)
        IF ABS(fTenNowN) < fZeroEpsN THEN
            _eState := eStSwitch;       (* 零位到位转切换步 / To switch *)
        ELSIF tonZero.Q THEN
            uCode := 16#003F;           (* 回零超时锁存故障（不无限等待）/ Latch the zeroing timeout *)
            _eState := eStIdle;         (* 回安全步 / Back to the safe step *)
        END_IF
    eStSwitch:                          (* 切换步：下发新配方参数并收周期 / Switch and close *)
        _bDone := TRUE;                 (* 完成脉冲置内部标志，段 3 输出 / Set internal done flag *)
        IF nCycles < DL_RCS_WRAP THEN
            nCycles := nCycles + 1;     (* 完成切换计数 / Count changeovers *)
        END_IF
        _eState := eStIdle;             (* 回空闲步 / Back to idle *)
ELSE
    _eState := eStIdle;                 (* ELSE 兜底回安全步 / ELSE fallback to safe step *)
END_CASE

(* === 段 3 · 输出映射与故障码（CASE 内未触碰输出枚举）=== *)
bSeqDone := _bDone;                     (* 完成脉冲输出（CASE 置位→此处映射）/ Done pulse mapped from internal flag *)
_bDone := FALSE;                        (* 单拍脉冲收口（置位与收口分离，防同拍抹除）/ One-scan pulse, no same-scan wipe *)
eStep := eStpIdle;                      (* 步映射默认 / Default mapping *)
IF _eState = eStValidate THEN
    eStep := eStpValidate;              (* 校验步映射 / Map validate *)
ELSIF _eState = eStTenZero THEN
    eStep := eStpTenZero;               (* 回零步映射 / Map zeroing *)
ELSIF _eState = eStSwitch THEN
    eStep := eStpSwitch;                (* 切换步映射 / Map switch *)
END_IF
bError := (uCode <> 16#0000);           (* 故障锁存回放 / Latched fault replay *)
uErrorId := WORD_TO_UDINT(uCode);       (* 码位单点写入（16#0000_003F 形态）/ Single write point *)
END_FUNCTION_BLOCK

(* ---- FB_DL_RollCompressForceBalance.st ---- *)
//==============================================================================
// 功能块：FB_DL_RollCompressForceBalance ｜ 中文名称：辊压机两侧轧制力平衡监视与液压纠偏
// 所属子库：DL_Process ｜ 版本：v1.0.0 ｜ 兼容：CODESYS V3.5+ / TwinCAT 3 / 汇川 InoProShop
// 功能描述：辊压机两侧轧制力差动平衡——压差 = 左力 - 右力，压差绝对值
//           超窗口（fDiffLimitKn）持续去抖窗 → 差动修调输出（液压比例
//           阀方向修调 fTrimPct，正 = 增左/减右向），修调带增益映射与
//           每拍限速（液压平稳性约束）；修调饱和（满幅）后压差仍持续
//           超窗 tSatTimeout → 判液压侧异常（纠偏能力耗尽），锁存故障；
//           压差回窗口内 → 修调按限速回零。压差进入窗口前给预警带信息
//           提示（供提前干预）。
// 遗留假设（R95 代理阈值三句）：① 代理值 = fCycleTimeS 组态扫描周期
//           [秒]（限速积分基量）；② 覆盖 0.001~0.1 秒任务周期范围；
//           ③ 覆盖不到的区间由调用方按实际任务周期重设该引脚负责，
//           该假设挂编译验证债。同拍多窗配比约束（R100）：
//           tSatTimeout > tDiffDebounce——饱和确认窗必须长于去抖窗，
//           否则压差尚未确认即误判饱和异常。
// 开源溯源 (Origin)：道莅原创实现（参考辊压机轧制力平衡与液压差动纠偏工程惯例 分类与参数域）
// 单位表：轧制力[千牛] / 压差[千牛] / 压差窗[千牛] / 修调[百分数] /
//         修调增益[百分数每千牛] / 限速[百分数每秒] / 时间[ms] / 扫描周期[秒]
// 错误码表：16#0005_01FC 信息级（压差进入预警带：超窗去抖计窗中，不置
//           bError）/ 16#0005_01FD 信息级（修调输出达限幅提示，不置
//           bError）/ 16#0005_033F 故障级（组态非法：压差窗/增益/限速/
//           周期域、时间窗 <= 0 或配比倒置（饱和窗 <= 去抖窗），或任一
//           输入非有限，置 bError）/ 16#0005_0340 故障级（压差持续超窗
//           且纠偏饱和：修调满幅后超窗持续 tSatTimeout，判液压侧异常
//           嫌疑，修调冻结，置 bError——该场景不可由 033F 的组态类判据
//           观测，属液压执行独立域）/ 16#0005_0341 故障级兜底（状态机
//           落 ELSE，置 bError 并撤修调）
// 状态机：E_DL_RollBalanceState（四态：eIdle=0 / eBalance=10 / eFrozen=20 /
//           eFault=99），CASE 含 ELSE 兜底，ELSE 置 0341 并撤修调
// 边界行为：① 组态非法 → 故障态锁存，bReset 复位；② 修调限速双向
//           （逼近与回零均限速，防液压冲击）；③ 修调饱和后压差回窗 →
//           正常回零路径（饱和不锁存，仅持续超窗才锁存故障）；④ 轧力
//           非有限 → 冻结修调安全侧（数据不可信不动液压）＋ 故障 033F
//           复用（R90：组态类「输入非法」语义扩覆盖）；⑤ 未使能修调
//           撤零并 bValid := FALSE；⑥ 安全侧 = 故障/冻结路径修调保持
//           进入时的值不再变化（液压跳变比保持更危险）。
// 修订历史：v1.0.0 2026-11-17 首版（R24 派单 · ROADMAP P1 §805）
//==============================================================================

(*------------------------------------------------------------------------------
 * 枚举: E_DL_RollBalanceState（归属本功能块，同文件发布，全库唯一定义）
 * 含义: 平衡监视相位，每个成员在 CASE 中有且仅有一个标签。
 *-----------------------------------------------------------------------------*)
TYPE E_DL_RollBalanceState :
(
    eIdle    := 0,   // 空闲：未使能 / Idle, not enabled
    eBalance := 10,  // 平衡：修调闭环运行 / Balance, trim loop running
    eFrozen  := 20,  // 冻结：纠偏饱和后持续超窗，修调保持 / Frozen, saturated trim held
    eFault   := 99   // 故障：组态非法/非有限/非法状态 / Fault, config, non-finite or illegal state
);
END_TYPE

FUNCTION_BLOCK FB_DL_RollCompressForceBalance
VAR_INPUT
    bEnable        : BOOL;                  // 平衡使能 [—] / Balance enable
    bReset         : BOOL;                  // 故障复位 [—]，上升沿清锁存 / Fault reset, rising edge clears latches
    fForceLeftKn   : LREAL;                 // 左侧轧制力 [千牛] / Left roll force [kN]
    fForceRightKn  : LREAL;                 // 右侧轧制力 [千牛] / Right roll force [kN]
    fDiffLimitKn   : LREAL := 10.0;         // 压差窗 [千牛]，须 > 0 / Differential window [kN]
    fTrimGainPctPerKn: LREAL := 1.0;        // 修调增益 [百分数每千牛] / Trim gain [percent/kN]
    fTrimRatePctS  : LREAL := 5.0;          // 修调限速 [百分数每秒]，须 > 0 / Trim slew rate [percent/s]
    fCycleTimeS    : LREAL := 0.01;         // 任务扫描周期 [秒]，须 > 0（R95 代理阈值） / Task scan cycle [s], must be > 0, R95 proxy
    tDiffDebounce  : TIME  := T#2S;         // 压差去抖窗 [ms]，须 > 0 / Differential debounce window [ms]
    tSatTimeout    : TIME  := T#30S;        // 饱和确认窗 [ms]，须 > 去抖窗（R100 配比） / Saturation confirm window [ms], must exceed the debounce
END_VAR
VAR_OUTPUT
    fTrimPct       : LREAL;                 // 差动修调输出 [百分数]，-100..100（正 = 增左向） / Differential trim output [percent], positive raises the left side
    bBalanceOk     : BOOL;                  // 压差在窗内 [—] / Differential inside the window
    bTrimSaturated : BOOL;                  // 修调饱和 [—] / Trim saturated
    eState         : E_DL_RollBalanceState; // 相位出口 [—] / Phase outlet
    eErr           : UDINT;                 // 错误码，0 = 无错，码位 16#0005_01FC 起信息级、16#0005_033F 起故障级（分带见错误码表） / Error code, 0 = no error, band info/fault per the code table
    bError         : BOOL;                  // 故障级标志，仅故障级错误置位 / Fault-class flag, set only on fault-level codes
    bValid         : BOOL;                  // 输出可用标志 / Outputs usable flag
END_VAR
VAR
    fbDebounce : TON;                       // 压差去抖计时（每拍无条件刷新）[ms] / Debounce timer, refreshed unconditionally
    fbSat      : TON;                       // 饱和确认计时（每拍无条件刷新）[ms] / Saturation confirm timer, refreshed unconditionally
    _eState    : E_DL_RollBalanceState := E_DL_RollBalanceState.eIdle; // 当前相位 / Current phase
    _bCfgBad   : BOOL;                      // 组态非法锁存 / Illegal config latch
    _bInfoOver : BOOL;                      // 预警信息当拍标志 / Over-window info flag of this scan
    _bInfoSat  : BOOL;                      // 限幅信息当拍标志 / Saturation info flag of this scan
    _fDiff     : LREAL;                     // 压差 [千牛] / Differential [kN]
    _fTrimTarget: LREAL;                    // 修调目标 [百分数] / Trim target [percent]
    _fStep     : LREAL;                     // 本拍限速步进 [百分数] / Per-scan slew step [percent]
    _bIllegal  : BOOL;                      // 非法状态标志 / Illegal state flag
    _bInit     : BOOL := FALSE;             // 首扫标志，初值 FALSE 取非判定 / First-scan flag, tested negated
END_VAR
VAR CONSTANT
    DL_RCF_INF      : LREAL := 1.7976931348623157E308; // LREAL 幅值上限 / LREAL magnitude ceiling
    DL_RCF_EPS      : LREAL := 1.0E-6;      // 浮点判零容差 [混合] / Float zero tolerance
    DL_RCF_TRIMMAX  : LREAL := 100.0;       // 修调满幅 [百分数] / Trim full scale [percent]
    DL_RCF_SAT_EPS  : LREAL := 0.5;         // 饱和判定容差 [百分数]（距满幅 0.5% 内判饱和） / Saturation tolerance [percent]
    DL_RCF_ZERO     : LREAL := 0.0;         // 零值常量，避免裸字面量 [混合] / Zero constant, avoids a bare literal
END_VAR

(*------------------------------------------------------------------------------
 * 段 1｜每拍预置：修调保持语义（预置不清零，冻结/故障须保持），标志预清零
 *      Trim kept by design (held in frozen and fault), flags pre-cleared
 *-----------------------------------------------------------------------------*)
bBalanceOk := FALSE;                     // 压差在窗电平先清（段 5 重置） / In-window level cleared first
bTrimSaturated := FALSE;                 // 饱和电平先清 / Saturated level cleared first
eErr   := 16#0000_0000;                  // 错误码每拍重算 / Error code recomputed
bError := FALSE;                         // 故障标志每拍重算 / Fault flag recomputed
bValid := FALSE;                         // 可用标志每拍重算 / Usable flag recomputed
_bInfoOver := FALSE;                     // 预警信息预清零 / Over-window info pre-cleared
_bInfoSat  := FALSE;                     // 限幅信息预清零 / Saturation info pre-cleared
_bIllegal  := FALSE;                     // 非法状态预清零 / Illegal flag pre-cleared

(*------------------------------------------------------------------------------
 * 段 2｜首扫初始化
 *      First-scan initialisation
 *-----------------------------------------------------------------------------*)
IF NOT _bInit THEN
    _eState  := E_DL_RollBalanceState.eIdle; // 相位空闲起步 / Phase starts idle
    _bCfgBad := FALSE;                   // 组态锁存清零 / Config latch cleared
    fTrimPct := DL_RCF_ZERO;             // 修调从零起步 / Trim starts at zero
    _bInit   := TRUE;                    // 首扫只做一次 / The first scan runs once
END_IF

(*------------------------------------------------------------------------------
 * 段 3｜组态防御闸：非有限（R79）+ 压差窗/增益/限速/周期/时间窗域（含 R100 配比）
 *      Configuration defense gates with the R100 ratio rule
 *-----------------------------------------------------------------------------*)
IF (fForceLeftKn <> fForceLeftKn) OR (ABS(fForceLeftKn) > DL_RCF_INF)
   OR (fForceRightKn <> fForceRightKn) OR (ABS(fForceRightKn) > DL_RCF_INF)
   OR (fDiffLimitKn <> fDiffLimitKn) OR (ABS(fDiffLimitKn) > DL_RCF_INF)
   OR (fTrimGainPctPerKn <> fTrimGainPctPerKn) OR (ABS(fTrimGainPctPerKn) > DL_RCF_INF)
   OR (fTrimRatePctS <> fTrimRatePctS) OR (ABS(fTrimRatePctS) > DL_RCF_INF)
   OR (fCycleTimeS <> fCycleTimeS) OR (ABS(fCycleTimeS) > DL_RCF_INF) THEN
    _bCfgBad := TRUE;                    // 非有限归组态非法锁存 / Non-finite folded into the config latch
END_IF
IF (NOT _bCfgBad) AND ((fDiffLimitKn <= DL_RCF_EPS) OR (fTrimRatePctS <= DL_RCF_EPS)
   OR (fCycleTimeS <= DL_RCF_EPS) OR (tDiffDebounce <= T#0MS)
   OR (tSatTimeout <= tDiffDebounce)) THEN
    _bCfgBad := TRUE;                    // 压差窗/限速/周期/时间窗域非法锁存（饱和窗须长于去抖窗） / Window domains latched, saturation window must exceed the debounce
END_IF
IF bReset THEN
    _bCfgBad := FALSE;                   // 复位清组态锁存 / Reset clears the config latch
END_IF

(*------------------------------------------------------------------------------
 * 段 4｜双计时无条件刷新（R40：CASE 之外每拍必调）
 *      Two timers refreshed unconditionally per R40
 *-----------------------------------------------------------------------------*)
fbDebounce(IN := (_eState = E_DL_RollBalanceState.eBalance)
                AND (ABS(_fDiff) > fDiffLimitKn), PT := tDiffDebounce); // 压差去抖窗 / Differential debounce window
fbSat(IN := (_eState = E_DL_RollBalanceState.eBalance)
           AND bTrimSaturated AND (ABS(_fDiff) > fDiffLimitKn), PT := tSatTimeout); // 饱和确认窗 / Saturation confirm window

(*------------------------------------------------------------------------------
 * 段 5｜相位机与修调链（CASE 含 ELSE 兜底；状态改写只出现在分支判据内，R39）
 *      Phase machine and the trim chain
 *-----------------------------------------------------------------------------*)
_fDiff := fForceLeftKn - fForceRightKn;  // 压差 [千牛] / Differential
CASE _eState OF

    E_DL_RollBalanceState.eIdle:           // 空闲：使能且组态合法进平衡态
        IF bEnable AND (NOT _bCfgBad) THEN
            _eState := E_DL_RollBalanceState.eBalance; // 进平衡 / To balance
        ELSIF bEnable AND _bCfgBad THEN
            _eState := E_DL_RollBalanceState.eFault; // 组态非法进故障 / Illegal config to fault
        END_IF

    E_DL_RollBalanceState.eBalance:        // 平衡：修调闭环 + 饱和确认
        IF (NOT bEnable) OR _bCfgBad THEN
            _eState := E_DL_RollBalanceState.eFault; // 异常转故障 / Anomaly, fault
        ELSE
            bBalanceOk := ABS(_fDiff) <= fDiffLimitKn; // 压差在窗电平 / In-window level
            _fTrimTarget := MIN(MAX(-fTrimGainPctPerKn * _fDiff,
                              -DL_RCF_TRIMMAX), DL_RCF_TRIMMAX); // 修调目标（负反馈向）双侧满幅钳位 / Trim target, both sides clamped
            _fStep := fTrimRatePctS * fCycleTimeS; // 本拍限速步进 [百分数] / Per-scan slew step
            fTrimPct := MIN(MAX(fTrimPct, _fTrimTarget - _fStep),
                            _fTrimTarget + _fStep); // 限速逼近目标（双向平稳） / Slew approach, smooth both ways
            fTrimPct := MIN(MAX(fTrimPct, -DL_RCF_TRIMMAX), DL_RCF_TRIMMAX); // 满幅终钳 / Final full-scale clamp
            bTrimSaturated := ABS(fTrimPct) >= (DL_RCF_TRIMMAX - DL_RCF_SAT_EPS); // 饱和判定 / Saturation verdict
            IF bTrimSaturated THEN
                _bInfoSat := TRUE;         // 修调达限幅提示（信息级） / Trim at limit, info
            ELSIF ABS(_fDiff) > fDiffLimitKn THEN
                _bInfoOver := TRUE;        // 压差超窗预警（去抖计窗中，信息级） / Over-window warning, info
            END_IF
            IF fbSat.Q THEN
                _eState := E_DL_RollBalanceState.eFrozen; // 饱和后持续超窗：修调冻结（拍 N 进入） / Saturated over-window, trim frozen
            END_IF
        END_IF

    E_DL_RollBalanceState.eFrozen:         // 冻结：修调保持进入时的值；压差回窗且复位后回平衡
        IF (NOT bEnable) OR _bCfgBad THEN
            _eState := E_DL_RollBalanceState.eFault; // 异常转故障 / Anomaly, fault
        ELSIF bReset AND (ABS(_fDiff) <= fDiffLimitKn) THEN
            _eState := E_DL_RollBalanceState.eBalance; // 复位且压差回窗回平衡 / Reset with the window back, to balance
        END_IF

    E_DL_RollBalanceState.eFault:          // 故障：复位沿且原因消失回平衡态
        IF bReset AND (NOT _bCfgBad) THEN
            _eState := E_DL_RollBalanceState.eBalance; // 回平衡 / Back to balance
        END_IF

    ELSE                                   // 非法状态兜底（R21：CASE 必带 ELSE）
        _bIllegal := TRUE;                 // 标记非法状态 / Flag the illegal state
        fTrimPct := DL_RCF_ZERO;           // 修调撤零（安全侧） / Trim cleared, safe side
        _eState := E_DL_RollBalanceState.eFault; // 回故障态 / Back to fault
END_CASE

(*------------------------------------------------------------------------------
 * 段 6｜码位出口与放行（故障级码 3 行内置 bError，R45/R101 配对）
 *      Code outlet and release, fault codes paired with bError
 *-----------------------------------------------------------------------------*)
IF _bIllegal THEN
    eErr   := 16#0005_0341;                // 故障级：状态机兜底 / Fault: state machine fallback
    bError := TRUE;                        // 置故障标志 / Raise the fault flag
ELSIF _bCfgBad THEN
    eErr   := 16#0005_033F;                // 故障级：组态非法 / Fault: illegal configuration
    bError := TRUE;                        // 置故障标志 / Raise the fault flag
ELSIF _eState = E_DL_RollBalanceState.eFrozen THEN
    eErr   := 16#0005_0340;                // 故障级：压差持续超窗且纠偏饱和 / Fault: sustained over-window with saturated trim
    bError := TRUE;                        // 置故障标志 / Raise the fault flag
ELSIF _bInfoSat THEN
    eErr := 16#0005_01FD;                  // 信息级：修调输出达限幅 / Info: trim at limit
ELSIF _bInfoOver THEN
    eErr := 16#0005_01FC;                  // 信息级：压差进入预警带 / Info: over-window warning
END_IF

IF (NOT bEnable) THEN
    fTrimPct := DL_RCF_ZERO;               // 未使能修调撤零（R72 显式路径） / Not enabled, trim to zero
END_IF
bValid := (NOT bError) AND bEnable AND (_eState <> E_DL_RollBalanceState.eIdle); // 空闲/故障/未使能输出不可用 / Outputs unusable in idle, fault or disabled
eState := _eState;                       // 相位出口 / Phase outlet
END_FUNCTION_BLOCK

(* ---- FB_DL_RollPressBitWord.st ---- *)
(*
  ==================================================================
  组件名 Component  : FB_DL_RollPressBitWord
  分类   Category   : DL_Process
  版本   Version    : 1.0.0
  功能   Purpose    : 辊压压力报警字位段打包。逐区（1..8）比较实测压力与逐区
                      高压阈 / 低压阈，带回差防抖，把报警状态打包为一个 16 位字：
                      低 8 位段 = 低压报警（位 i-1 对应区 i），
                      高 8 位段 = 高压报警（位 8+i-1 对应区 i），
                      另出无效区掩码字（该区不可判：阈值非法或压力非有限）。
  溯源   Origin     : 逐区位段打包与回差防抖为通用报警字组织方式；本件为 clean-room
                      实现，仅借鉴来源分类与参数域组织（来源标签 roadmap-p2-rollpress），
                      道莅原创设计，未复制任何闭源代码行。
  平台   Platform   : 纯 IEC 61131-3（WORD / SHL / NOT / AND / OR，无私有库）
  作者   Author     : 道莅代码库 · PLC 编程专家（R55）
  ------------------------------------------------------------------
  边界 Boundary     :
                      一 本件只做压力报警字打包，不驱动辊缝、不做停机决策（属主边界）；
                      二 回差判据挂在报警字自身状态上（已置位者按 阈 - 回差 复位）；
                      三 非有限压力不判高低压，只置无效位，出口报警位保持上拍；
                      四 阈值非法（高阈不高于低阈或非有限）→ 该区无效 + 故障锁存；
                      五 无全局变量、无外部变量声明、无物理地址寻址。
  输出契约 Output contract:
                      wAlarmWord 低字节为低压段、高字节为高压段，两段互不跨用；
                      自证向量：仅 1 区低压 → 16#0001，仅 1 区高压 → 16#0100，
                      1 区低压且 8 区高压 → 16#0180；
                      nFirstAlarmZone 为 1..8，无报警为 0；uAlarmCount 为本拍置位数；
                      eCause 故障级成因与 bError 配对（R45），信息级永不置 bError。
  修订记录 Revision  :
    2026-11-20  v1.0.0  R55 首版（批 1 · 序号 5）
  ==================================================================
*)

TYPE E_DL_RpbCause :
(
    eNone       := 0,   // 无成因 / no cause
    eThrBad     := 1,   // 阈值非法：高阈不高于低阈或非有限（故障级，与 bError 配对）/ illegal threshold, high not above low or non-finite, a fault paired with bError
    eCountBad   := 2,   // 区数越域已回钳（信息级）/ zone count out of domain and clamped, informational
    ePressBad   := 3    // 压力非有限，该区不可判（信息级）/ non-finite pressure, the zone is undecidable, informational
);
END_TYPE

FUNCTION_BLOCK FB_DL_RollPressBitWord
VAR_INPUT
    bEnable      : BOOL := TRUE;             // 使能，失能时报警字冻结保持末值 [-] / enable, the alarm word freezes and holds its last value when disabled
    bReset       : BOOL := FALSE;           // 复位上升沿清报警位与故障锁存 [-] / reset rising edge clears the alarm bits and the fault latch
    nZoneCount   : INT := 8;                 // 参与判定的区数 [个]，域 1..8 / participating zones [count], domain 1 to 8
    fHystBar     : REAL := 0.5;              // 回差带 [巴]，域 大于等于零 / hysteresis band [bar], domain zero and above
END_VAR
VAR_IN_OUT
    afPressBar   : ARRAY[1..8] OF REAL;      // 逐区压力实测 [巴]，引用型入参由调用方持有 / per zone measured pressure [bar], reference parameter owned by the caller
    afPressHiBar : ARRAY[1..8] OF REAL;      // 逐区高压报警阈 [巴]，引用型入参由调用方持有 / per zone high alarm threshold [bar], reference parameter owned by the caller
    afPressLoBar : ARRAY[1..8] OF REAL;      // 逐区低压报警阈 [巴]，引用型入参由调用方持有 / per zone low alarm threshold [bar], reference parameter owned by the caller
END_VAR
VAR_OUTPUT
    wAlarmWord   : WORD := 16#0000;          // 打包报警字：低字节低压段 / 高字节高压段 [-] / packed alarm word, low byte for the low segment and high byte for the high segment
    wLowWord     : WORD := 16#0000;          // 低压报警段（位 i-1 对应区 i）[-] / low pressure alarm segment, bit i minus one maps to zone i
    wHighWord    : WORD := 16#0000;          // 高压报警段（位 i-1 对应区 i）[-] / high pressure alarm segment, bit i minus one maps to zone i
    wInvalidWord : WORD := 16#0000;          // 无效区掩码（不可判的区）[-] / invalid zone mask for undecidable zones
    bAnyAlarm    : BOOL := FALSE;            // 任一报警置位 [-] / any alarm bit set
    nFirstAlarmZone : INT := 0;              // 首个报警区号 [区号]，无报警为 0 / first alarming zone number, zero when none
    uAlarmCount  : UINT := 0;                // 本拍报警位数 [位] / number of alarm bits this scan
    eCause       : E_DL_RpbCause := E_DL_RpbCause.eNone; // 成因出口 [枚举] / cause outlet [enum]
    bError       : BOOL := FALSE;            // 故障锁存标志 [-] / fault latch flag
END_VAR
VAR
    rtReset      : R_TRIG;                   // 复位沿检测，段 0 无条件刷新 / reset edge detector, refreshed unconditionally in segment zero
    _eCause      : E_DL_RpbCause := E_DL_RpbCause.eNone; // 内部成因，故障级锁存、信息级每拍重算 / internal cause, latched for faults and recomputed for information
    _bFault      : BOOL := FALSE;            // 故障锁存位（阈值非法）/ fault latch bit for an illegal threshold
    _bInit       : BOOL := FALSE;            // 首扫初始化完成标志（R310）/ first scan initialisation flag
    _bAnyAlarm   : BOOL := FALSE;            // 任一报警标志工作值（出口映射源）[-] / any-alarm working flag, source of the outlet
    _bZoneBad    : BOOL := FALSE;            // 本区不可判（阈值非法或压力非有限）[-] / the zone is undecidable
    _bPressOk    : BOOL := FALSE;            // 本区压力有限 [-] / the zone pressure is finite
    _bThrOk      : BOOL := FALSE;            // 本区阈值合法 [-] / the zone thresholds are legal
    _bPressNonFin: BOOL := FALSE;            // 本拍出现非有限压力 [-] / a non-finite pressure occurred this scan
    _bCountClamped : BOOL := FALSE;          // 区数被回钳 [-] / the zone count was clamped
    _bHiBit      : BOOL := FALSE;            // 本区高压报警位当前值 [-] / current high alarm bit of the zone
    _bLoBit      : BOOL := FALSE;            // 本区低压报警位当前值 [-] / current low alarm bit of the zone
    _nUseCount   : INT := 0;                 // 钳定后的区数 [个] / clamped zone count
    _nIdx        : INT := 0;                 // 区游标（1 起，回钳 1..8）[区号] / zone cursor, one-based, clamped one through eight
    _fPress      : REAL := 0.0;              // 本区压力暂存 [巴] / zone pressure held in a local [bar]
    _fHi         : REAL := 0.0;              // 本区高压阈暂存 [巴] / zone high threshold held in a local [bar]
    _fLo         : REAL := 0.0;              // 本区低压阈暂存 [巴] / zone low threshold held in a local [bar]
    _fHiReset    : REAL := 0.0;              // 高压回差复位点 [巴] / high hysteresis reset point [bar]
    _fLoReset    : REAL := 0.0;              // 低压回差复位点 [巴] / low hysteresis reset point [bar]
    _fHyst       : REAL := 0.0;              // 钳定后的回差 [巴] / clamped hysteresis [bar]
    _wLo         : WORD := 16#0000;          // 低压段工作字，兼作回差状态 / low segment working word, also the hysteresis state
    _wHi         : WORD := 16#0000;          // 高压段工作字，兼作回差状态 / high segment working word, also the hysteresis state
    _wInv        : WORD := 16#0000;          // 无效区工作字 / invalid zone working word
    _wBit        : WORD := 16#0001;          // 本区位掩码，先移位后置位（R327）/ zone bit mask, shift before setting
END_VAR
VAR CONSTANT
    DL_RPB_MAX      : INT := 8;              // 区容量与游标回钳上界 [个] / zone capacity and cursor clamp upper bound
    DL_RPB_SEG_SHIFT: INT := 8;              // 高压段移入高字节的位移量 [位]，常量 8 小于字宽 16 / shift moving the high segment into the high byte, the constant eight is below the word width sixteen
    DL_RPB_MASK_NONE: WORD := 16#0000;       // 空掩码常量 [-] / empty mask constant
    DL_RPB_MASK_ONE : WORD := 16#0001;       // 单位位常量 [-] / single bit constant
    DL_RPB_HYST_MAX : REAL := 100.0;         // 回差上限 [巴]，防回差吞掉整个量程 / hysteresis ceiling against swallowing the whole range [bar]
    DL_RPB_PRESS_MAX: REAL := 1.0E6;         // 压力量级上限，防量纲错配 [巴] / pressure magnitude ceiling against a dimension mismatch [bar]
END_VAR

// 段 0｜复位沿无条件周期刷新（禁入分支）/ segment 0, unconditional refresh of the reset edge, never inside a branch
rtReset(CLK := bReset); // 复位沿无条件刷新 / unconditional refresh of the reset edge

// 段 1｜首扫初始化（R310）/ segment 1, first scan initialisation
IF NOT _bInit THEN // 首扫一拍 / the very first scan
    _bInit := TRUE; // 置首扫完成标志 / raise the first scan flag
    _bFault := FALSE; // 故障锁存清零 / clear the fault latch
    _eCause := E_DL_RpbCause.eNone; // 成因清零 / clear the cause
    _wLo := DL_RPB_MASK_NONE; // 低压段清零 / clear the low segment
    _wHi := DL_RPB_MASK_NONE; // 高压段清零 / clear the high segment
    _wInv := DL_RPB_MASK_NONE; // 无效字清零 / clear the invalid word
END_IF

// 段 2｜复位沿作用域：清报警位 / 清无效字 / 清故障锁存（三项逐项声明）/ segment 2, reset edge scope declared item by item
IF rtReset.Q THEN // 复位沿 / reset edge
    _bFault := FALSE; // 作用域一：清故障锁存 / scope one, clear the fault latch
    _eCause := E_DL_RpbCause.eNone; // 作用域一：清成因 / scope one, clear the cause
    _wLo := DL_RPB_MASK_NONE; // 作用域二：清低压报警位 / scope two, clear the low alarm bits
    _wHi := DL_RPB_MASK_NONE; // 作用域二：清高压报警位 / scope two, clear the high alarm bits
    _wInv := DL_RPB_MASK_NONE; // 作用域三：清无效字 / scope three, clear the invalid word
END_IF

// 段 3｜区数回钳与回差域闸 / segment 3, zone count clamping and hysteresis domain gate
_bCountClamped := FALSE; // 回钳标志预置假 / preset the clamp flag to false
_nUseCount := nZoneCount; // 区数直通 / zone count passes through
IF _nUseCount < 1 THEN // 下越界 / below the lower bound
    _nUseCount := 1; // 回钳到 1 / clamp to one
    _bCountClamped := TRUE; // 置回钳标志 / raise the clamp flag
ELSIF _nUseCount > DL_RPB_MAX THEN // 上越界 / above the upper bound
    _nUseCount := DL_RPB_MAX; // 回钳到容量上限 / clamp to the capacity ceiling
    _bCountClamped := TRUE; // 置回钳标志 / raise the clamp flag
END_IF
_fHyst := fHystBar; // 回差直通 / hysteresis passes through
IF (_fHyst <> _fHyst) OR ((_fHyst - _fHyst) <> (_fHyst - _fHyst)) THEN // 回差非有限 / hysteresis non-finite
    _fHyst := 0.0; // 非有限归零（等价无回差）/ zeroed, equivalent to no hysteresis
END_IF
IF _fHyst < 0.0 THEN // 回差为负 / hysteresis negative
    _fHyst := 0.0; // 钳零 / clamped to zero
ELSIF _fHyst > DL_RPB_HYST_MAX THEN // 回差过大 / hysteresis too large
    _fHyst := DL_RPB_HYST_MAX; // 钳到上限 / clamped to the ceiling
END_IF
IF NOT bEnable THEN // 失能：报警字冻结保持末值（R191 显式声明）/ disabled, the alarm word freezes and holds its last value
    _nUseCount := 0; // 区数置零使主循环不执行 / the zone count is zeroed so the main loop does not run
END_IF

// 段 4｜逐区判定主循环：阈值闸 → 压力闸 → 回差判据 → 位打包（先移位后置位）/ segment 4, per zone loop with threshold gate, pressure gate, hysteresis criterion and bit packing
_bPressNonFin := FALSE; // 非有限压力标志清零 / clear the non-finite pressure flag
_nIdx := 1; // 游标自 1 起，上界由 _nUseCount 约束 / the cursor starts at one, bounded by the usable count
WHILE _nIdx <= _nUseCount DO // 循环上界为钳定后的区数，天然不越 8 / the loop bound is the clamped count, never beyond eight
    _wBit := SHL(DL_RPB_MASK_ONE, _nIdx - 1); // 本区位掩码，位移量 0..7 由数组边界与循环上界共同证明 / zone bit mask, the shift zero through seven is proven by the array and loop bounds
    _fPress := afPressBar[_nIdx]; // 压力暂存 / pressure held in a local
    _fHi := afPressHiBar[_nIdx]; // 高压阈暂存 / high threshold held in a local
    _fLo := afPressLoBar[_nIdx]; // 低压阈暂存 / low threshold held in a local
    _bThrOk := (_fHi = _fHi) AND ((_fHi - _fHi) = (_fHi - _fHi)) AND (_fLo = _fLo) AND ((_fLo - _fLo) = (_fLo - _fLo)) AND (_fHi > _fLo); // 阈值有限且高阈高于低阈 / thresholds finite with the high above the low
    _bPressOk := (_fPress = _fPress) AND ((_fPress - _fPress) = (_fPress - _fPress)) AND (ABS(_fPress) <= DL_RPB_PRESS_MAX); // 压力有限且量级可信 / pressure finite with a credible magnitude
    _bZoneBad := FALSE; // 本区不可判标志预置假 / preset the undecidable flag to false
    IF NOT _bThrOk THEN // 阈值非法 / illegal threshold
        _bZoneBad := TRUE; // 本区不可判 / the zone is undecidable
        IF NOT _bFault THEN // 未锁存才记故障 / record the fault only when not yet latched
            _bFault := TRUE; // 置故障锁存 / raise the fault latch
            _eCause := E_DL_RpbCause.eThrBad; // 故障级成因 (R45 配对 bError) / fault grade cause paired with bError
        END_IF
    ELSIF NOT _bPressOk THEN // 压力非有限 / pressure non-finite
        _bZoneBad := TRUE; // 本区不可判 / the zone is undecidable
        _bPressNonFin := TRUE; // 记非有限压力成因 / record the non-finite pressure cause
    END_IF
    _wInv := _wInv AND NOT _wBit; // 先假定本区可判，清无效位 / assume the zone is decidable and clear the invalid bit
    IF _bZoneBad THEN // 本区不可判 / the zone is undecidable
        _wInv := _wInv OR _wBit; // 置无效位 / set the invalid bit
        _wLo := _wLo AND NOT _wBit; // 低压位保持清零（不可判不报警）/ the low bit stays cleared, nothing is decided
        _wHi := _wHi AND NOT _wBit; // 高压位保持清零（不可判不报警）/ the high bit stays cleared, nothing is decided
    ELSE
        _bLoBit := ((_wLo AND _wBit) <> DL_RPB_MASK_NONE); // 低压位当前值 / current low bit
        _bHiBit := ((_wHi AND _wBit) <> DL_RPB_MASK_NONE); // 高压位当前值 / current high bit
        _fLoReset := _fLo + _fHyst; // 低压回差复位点（已报警者高于此值才复位）/ low hysteresis reset point
        _fHiReset := _fHi - _fHyst; // 高压回差复位点（已报警者低于此值才复位）/ high hysteresis reset point
        IF _bLoBit THEN // 低压已报警 / the low alarm is active
            IF _fPress > _fLoReset THEN // 回升越过回差复位点 / recovered above the reset point
                _wLo := _wLo AND NOT _wBit; // 复位低压位 / clear the low bit
            END_IF
        ELSE // 低压未报警 / the low alarm is inactive
            IF _fPress < _fLo THEN // 低于低压阈 / below the low threshold
                _wLo := _wLo OR _wBit; // 置低压位 / set the low bit
            END_IF
        END_IF
        IF _bHiBit THEN // 高压已报警 / the high alarm is active
            IF _fPress < _fHiReset THEN // 回落越过回差复位点 / recovered below the reset point
                _wHi := _wHi AND NOT _wBit; // 复位高压位 / clear the high bit
            END_IF
        ELSE // 高压未报警 / the high alarm is inactive
            IF _fPress > _fHi THEN // 高于高压阈 / above the high threshold
                _wHi := _wHi OR _wBit; // 置高压位 / set the high bit
            END_IF
        END_IF
    END_IF
    _nIdx := _nIdx + 1; // 游标递增 / increment the cursor
END_WHILE

// 段 5｜字位段打包：低字节放低压段、高字节放高压段，两段互不跨用 / segment 5, segment packing with the low byte for the low segment and the high byte for the high segment
wLowWord := _wLo; // 低压段出口 / low segment outlet
wHighWord := _wHi; // 高压段出口 / high segment outlet
wInvalidWord := _wInv; // 无效区掩码出口 / invalid zone mask outlet
wAlarmWord := _wLo OR SHL(_wHi, DL_RPB_SEG_SHIFT); // 两段合成，位移量为常量八 / both segments combined with the constant shift of eight

// 段 6｜统计：报警位数与首个报警区号（自 1 区起顺序扫，命中即止）/ segment 6, statistics for the alarm count and the first alarming zone
_bAnyAlarm := FALSE; // 任一报警标志预置假 / preset the any alarm flag to false
uAlarmCount := 0; // 报警位数清零 / clear the alarm bit count
nFirstAlarmZone := 0; // 首个报警区号清零 / clear the first alarming zone
_nIdx := 1; // 游标自 1 起 / the cursor starts at one
WHILE _nIdx <= DL_RPB_MAX DO // 全容量扫查，未参与区恒为零位 / sweep the full capacity because unused zones stay cleared
    _wBit := SHL(DL_RPB_MASK_ONE, _nIdx - 1); // 本区位掩码 / zone bit mask
    IF ((_wLo AND _wBit) <> DL_RPB_MASK_NONE) OR ((_wHi AND _wBit) <> DL_RPB_MASK_NONE) THEN // 本区任一报警位 / any alarm bit of this zone
        _bAnyAlarm := TRUE; // 置任一报警标志 / raise the any alarm flag
        uAlarmCount := uAlarmCount + 1; // 报警位数递增 / increment the alarm count
        IF nFirstAlarmZone = 0 THEN // 尚未记录首个 / nothing recorded yet
            nFirstAlarmZone := _nIdx; // 记录首个报警区号 / record the first alarming zone
        END_IF
    END_IF
    _nIdx := _nIdx + 1; // 游标递增 / increment the cursor
END_WHILE
bAnyAlarm := _bAnyAlarm; // 任一报警出口（挂状态量，非单拍标志）/ any alarm outlet, a state quantity

// 段 7｜成因分派（固定优先级：故障 > 回钳 > 非有限压力 > 无成因）/ segment 7, cause dispatch with a fixed priority
IF _bFault THEN // 故障锁存优先 / the fault latch takes priority
    _eCause := E_DL_RpbCause.eThrBad; // 故障级成因锁存回放 / the fault cause is replayed from the latch
ELSIF _bCountClamped THEN // 区数被回钳 / the zone count was clamped
    _eCause := E_DL_RpbCause.eCountBad; // 信息级成因 / informational cause
ELSIF _bPressNonFin THEN // 存在非有限压力 / a non-finite pressure occurred
    _eCause := E_DL_RpbCause.ePressBad; // 信息级成因 / informational cause
ELSE
    _eCause := E_DL_RpbCause.eNone; // 无成因 / no cause
END_IF

// 段 8｜统一出口 / segment 8, unified outlet
eCause := _eCause; // 成因出口单点映射 / single-point cause outlet mapping
bError := _bFault; // 故障标志与锁存位同源 / the fault flag shares the latch source
END_FUNCTION_BLOCK
